  movel([0.337067, -0.792207, -2.792280, -1.127903, 1.570796, 1.907863],accel_mss,speed_ms,0,blend_radius_m)
  movel([0.336030, -0.792065, -2.792303, -1.128021, 1.570796, 1.906826],accel_mss,speed_ms,0,blend_radius_m)
  movel([0.330509, -0.790300, -2.792596, -1.129493, 1.570796, 1.901306],accel_mss,speed_ms,0,blend_radius_m)
  movel([0.325271, -0.788116, -2.792957, -1.131316, 1.570796, 1.896067],accel_mss,speed_ms,0,blend_radius_m)
  movel([0.320318, -0.785517, -2.793383, -1.133490, 1.570796, 1.891115],accel_mss,speed_ms,0,blend_radius_m)
  movel([0.315671, -0.782494, -2.793873, -1.136022, 1.570796, 1.886468],accel_mss,speed_ms,0,blend_radius_m)
  movel([0.314088, -0.781197, -2.794083, -1.137109, 1.570796, 1.884885],accel_mss,speed_ms,0,blend_radius_m)
  movel([0.312919, -0.779429, -2.794366, -1.138594, 1.570796, 1.883716],accel_mss,speed_ms,0,blend_radius_m)
  movel([0.312565, -0.778043, -2.794588, -1.139758, 1.570796, 1.883362],accel_mss,speed_ms,0,blend_radius_m)
  movel([0.312427, -0.776467, -2.794838, -1.141084, 1.570796, 1.883224],accel_mss,speed_ms,0,blend_radius_m)
  movel([0.312533, -0.772984, -2.795388, -1.144017, 1.570796, 1.883329],accel_mss,speed_ms,0,blend_radius_m)
  movel([0.314201, -0.759545, -2.797451, -1.155393, 1.570796, 1.884998],accel_mss,speed_ms,0,blend_radius_m)
  movel([0.314322, -0.755972, -2.797984, -1.158433, 1.570796, 1.885118],accel_mss,speed_ms,0,blend_radius_m)
  movel([0.313995, -0.753066, -2.798414, -1.160909, 1.570796, 1.884791],accel_mss,speed_ms,0,blend_radius_m)
  movel([0.313608, -0.751988, -2.798572, -1.161829, 1.570796, 1.884404],accel_mss,speed_ms,0,blend_radius_m)
  movel([0.313044, -0.751216, -2.798685, -1.162488, 1.570796, 1.883841],accel_mss,speed_ms,0,blend_radius_m)
  movel([0.312284, -0.750809, -2.798744, -1.162836, 1.570796, 1.883080],accel_mss,speed_ms,0,blend_radius_m)
  movel([0.311307, -0.750804, -2.798745, -1.162840, 1.570796, 1.882104],accel_mss,speed_ms,0,blend_radius_m)
  movel([0.309324, -0.751441, -2.798652, -1.162296, 1.570796, 1.880120],accel_mss,speed_ms,0,blend_radius_m)
  movel([0.308425, -0.751616, -2.798626, -1.162147, 1.570796, 1.879221],accel_mss,speed_ms,0,blend_radius_m)
  movel([0.307786, -0.751386, -2.798660, -1.162343, 1.570796, 1.878582],accel_mss,speed_ms,0,blend_radius_m)
  movel([0.307584, -0.750201, -2.798833, -1.163355, 1.570796, 1.878380],accel_mss,speed_ms,0,blend_radius_m)
  movel([0.307977, -0.748520, -2.799077, -1.164791, 1.570796, 1.878773],accel_mss,speed_ms,0,blend_radius_m)
  movel([0.309463, -0.743009, -2.799868, -1.169512, 1.570796, 1.880260],accel_mss,speed_ms,0,blend_radius_m)
  movel([0.310630, -0.737685, -2.800619, -1.174085, 1.570796, 1.881426],accel_mss,speed_ms,0,blend_radius_m)
  movel([0.312165, -0.727491, -2.802019, -1.182879, 1.570796, 1.882961],accel_mss,speed_ms,0,blend_radius_m)
  movel([0.312944, -0.717680, -2.803320, -1.191389, 1.570796, 1.883740],accel_mss,speed_ms,0,blend_radius_m)
  movel([0.313326, -0.707992, -2.804562, -1.199834, 1.570796, 1.884122],accel_mss,speed_ms,0,blend_radius_m)
  speed_ms = 0.005
  movel([0.313326, -0.701025, -2.797945, -1.213418, 1.570796, 1.884122],accel_mss,speed_ms,0,blend_radius_m)
  speed_ms = 0.040
  movel([0.305588, -0.719229, -2.795588, -1.197572, 1.570796, 1.876385],accel_mss,speed_ms,0,blend_radius_m)
  speed_ms = 0.005
  movel([0.305588, -0.726439, -2.802160, -1.183790, 1.570796, 1.876385],accel_mss,speed_ms,0,blend_radius_m)
  speed_ms = 0.025
  movel([0.301170, -0.738509, -2.800504, -1.173377, 1.570796, 1.871966],accel_mss,speed_ms,0,blend_radius_m)
  movel([0.298692, -0.744594, -2.799642, -1.168153, 1.570796, 1.869489],accel_mss,speed_ms,0,blend_radius_m)
  movel([0.296052, -0.750689, -2.798762, -1.162938, 1.570796, 1.866849],accel_mss,speed_ms,0,blend_radius_m)
  movel([0.293909, -0.749383, -2.798952, -1.164054, 1.570796, 1.864706],accel_mss,speed_ms,0,blend_radius_m)
  movel([0.293492, -0.749233, -2.798974, -1.164182, 1.570796, 1.864289],accel_mss,speed_ms,0,blend_radius_m)
  movel([0.292925, -0.749435, -2.798944, -1.164009, 1.570796, 1.863721],accel_mss,speed_ms,0,blend_radius_m)
  movel([0.292315, -0.750102, -2.798847, -1.163439, 1.570796, 1.863111],accel_mss,speed_ms,0,blend_radius_m)
  movel([0.291839, -0.750915, -2.798729, -1.162745, 1.570796, 1.862635],accel_mss,speed_ms,0,blend_radius_m)
  movel([0.288894, -0.755925, -2.797991, -1.158473, 1.570796, 1.859691],accel_mss,speed_ms,0,blend_radius_m)
  movel([0.285493, -0.760805, -2.797261, -1.154323, 1.570796, 1.856290],accel_mss,speed_ms,0,blend_radius_m)
  movel([0.284595, -0.761864, -2.797101, -1.153424, 1.570796, 1.855391],accel_mss,speed_ms,0,blend_radius_m)
  movel([0.283710, -0.762451, -2.797012, -1.152926, 1.570796, 1.854506],accel_mss,speed_ms,0,blend_radius_m)
  movel([0.283279, -0.762203, -2.797050, -1.153136, 1.570796, 1.854075],accel_mss,speed_ms,0,blend_radius_m)
  movel([0.283199, -0.761526, -2.797152, -1.153711, 1.570796, 1.853995],accel_mss,speed_ms,0,blend_radius_m)
  movel([0.283611, -0.756734, -2.797871, -1.157784, 1.570796, 1.854408],accel_mss,speed_ms,0,blend_radius_m)
  movel([0.284807, -0.751427, -2.798654, -1.162308, 1.570796, 1.855604],accel_mss,speed_ms,0,blend_radius_m)
  speed_ms = 0.005
  movel([0.284807, -0.743907, -2.792145, -1.176337, 1.570796, 1.855604],accel_mss,speed_ms,0,blend_radius_m)
  speed_ms = 0.040
  movel([0.290706, -0.750918, -2.791114, -1.170358, 1.570796, 1.861503],accel_mss,speed_ms,0,blend_radius_m)
  speed_ms = 0.005
  movel([0.290706, -0.758522, -2.797604, -1.156263, 1.570796, 1.861503],accel_mss,speed_ms,0,blend_radius_m)
  speed_ms = 0.025
  movel([0.289009, -0.766268, -2.796430, -1.149691, 1.570796, 1.859805],accel_mss,speed_ms,0,blend_radius_m)
  movel([0.287811, -0.770306, -2.795806, -1.146277, 1.570796, 1.858608],accel_mss,speed_ms,0,blend_radius_m)
  movel([0.284778, -0.778595, -2.794500, -1.139294, 1.570796, 1.855575],accel_mss,speed_ms,0,blend_radius_m)
  movel([0.282956, -0.782810, -2.793822, -1.135757, 1.570796, 1.853753],accel_mss,speed_ms,0,blend_radius_m)
  movel([0.278747, -0.791286, -2.792433, -1.128671, 1.570796, 1.849544],accel_mss,speed_ms,0,blend_radius_m)
  movel([0.279478, -0.788663, -2.792867, -1.130860, 1.570796, 1.850275],accel_mss,speed_ms,0,blend_radius_m)
  movel([0.279565, -0.786419, -2.793235, -1.132735, 1.570796, 1.850361],accel_mss,speed_ms,0,blend_radius_m)
  movel([0.279016, -0.784705, -2.793515, -1.134169, 1.570796, 1.849813],accel_mss,speed_ms,0,blend_radius_m)
  movel([0.277841, -0.783676, -2.793682, -1.135031, 1.570796, 1.848637],accel_mss,speed_ms,0,blend_radius_m)
  speed_ms = 0.005
  movel([0.277841, -0.775786, -2.787260, -1.149343, 1.570796, 1.848637],accel_mss,speed_ms,0,blend_radius_m)
  speed_ms = 0.040
  movel([0.251919, -0.792770, -2.784449, -1.135169, 1.570796, 1.822716],accel_mss,speed_ms,0,blend_radius_m)
  speed_ms = 0.005
  movel([0.251919, -0.800843, -2.790822, -1.120725, 1.570796, 1.822716],accel_mss,speed_ms,0,blend_radius_m)
  speed_ms = 0.025
  movel([0.247378, -0.806648, -2.789820, -1.115921, 1.570796, 1.818174],accel_mss,speed_ms,0,blend_radius_m)
  movel([0.242549, -0.812092, -2.788864, -1.111433, 1.570796, 1.813345],accel_mss,speed_ms,0,blend_radius_m)
  movel([0.237519, -0.817097, -2.787971, -1.107321, 1.570796, 1.808315],accel_mss,speed_ms,0,blend_radius_m)
  movel([0.232368, -0.821580, -2.787160, -1.103649, 1.570796, 1.803164],accel_mss,speed_ms,0,blend_radius_m)
  movel([0.233688, -0.818996, -2.787629, -1.105764, 1.570796, 1.804484],accel_mss,speed_ms,0,blend_radius_m)
  movel([0.234683, -0.816593, -2.788062, -1.107734, 1.570796, 1.805479],accel_mss,speed_ms,0,blend_radius_m)
  movel([0.235280, -0.814585, -2.788421, -1.109383, 1.570796, 1.806076],accel_mss,speed_ms,0,blend_radius_m)
  movel([0.235407, -0.813183, -2.788670, -1.110536, 1.570796, 1.806203],accel_mss,speed_ms,0,blend_radius_m)
  movel([0.234984, -0.812617, -2.788771, -1.111001, 1.570796, 1.805780],accel_mss,speed_ms,0,blend_radius_m)
  movel([0.234547, -0.812711, -2.788754, -1.110924, 1.570796, 1.805344],accel_mss,speed_ms,0,blend_radius_m)
  movel([0.233940, -0.813094, -2.788686, -1.110609, 1.570796, 1.804736],accel_mss,speed_ms,0,blend_radius_m)
  movel([0.232209, -0.814833, -2.788377, -1.109180, 1.570796, 1.803005],accel_mss,speed_ms,0,blend_radius_m)
  movel([0.227802, -0.820578, -2.787342, -1.104469, 1.570796, 1.798598],accel_mss,speed_ms,0,blend_radius_m)
  movel([0.225752, -0.823067, -2.786889, -1.102433, 1.570796, 1.796549],accel_mss,speed_ms,0,blend_radius_m)
  movel([0.221376, -0.827745, -2.786027, -1.098617, 1.570796, 1.792172],accel_mss,speed_ms,0,blend_radius_m)
  movel([0.219102, -0.829874, -2.785631, -1.096884, 1.570796, 1.789898],accel_mss,speed_ms,0,blend_radius_m)
  movel([0.216804, -0.831814, -2.785268, -1.095307, 1.570796, 1.787600],accel_mss,speed_ms,0,blend_radius_m)
  movel([0.214506, -0.833546, -2.784942, -1.093901, 1.570796, 1.785302],accel_mss,speed_ms,0,blend_radius_m)
  movel([0.212240, -0.835024, -2.784662, -1.092702, 1.570796, 1.783037],accel_mss,speed_ms,0,blend_radius_m)
  movel([0.215104, -0.830931, -2.785433, -1.096025, 1.570796, 1.785901],accel_mss,speed_ms,0,blend_radius_m)
  movel([0.217906, -0.826781, -2.786206, -1.099402, 1.570796, 1.788702],accel_mss,speed_ms,0,blend_radius_m)
  movel([0.219209, -0.824080, -2.786703, -1.101606, 1.570796, 1.790005],accel_mss,speed_ms,0,blend_radius_m)
  movel([0.219966, -0.821533, -2.787169, -1.103687, 1.570796, 1.790763],accel_mss,speed_ms,0,blend_radius_m)
  movel([0.219920, -0.820731, -2.787315, -1.104343, 1.570796, 1.790716],accel_mss,speed_ms,0,blend_radius_m)
  movel([0.219466, -0.820469, -2.787362, -1.104558, 1.570796, 1.790262],accel_mss,speed_ms,0,blend_radius_m)
  movel([0.218525, -0.820910, -2.787282, -1.104197, 1.570796, 1.789321],accel_mss,speed_ms,0,blend_radius_m)
  movel([0.217006, -0.822224, -2.787043, -1.103122, 1.570796, 1.787803],accel_mss,speed_ms,0,blend_radius_m)
  movel([0.209003, -0.830286, -2.785554, -1.096549, 1.570796, 1.779799],accel_mss,speed_ms,0,blend_radius_m)
  movel([0.205006, -0.833828, -2.784889, -1.093672, 1.570796, 1.775803],accel_mss,speed_ms,0,blend_radius_m)
  movel([0.203015, -0.835288, -2.784612, -1.092488, 1.570796, 1.773811],accel_mss,speed_ms,0,blend_radius_m)
  movel([0.201023, -0.836475, -2.784387, -1.091527, 1.570796, 1.771819],accel_mss,speed_ms,0,blend_radius_m)
  speed_ms = 0.005
  movel([0.201023, -0.828056, -2.778123, -1.106210, 1.570796, 1.771819],accel_mss,speed_ms,0,blend_radius_m)
  speed_ms = 0.040
  movel([0.238662, -0.773617, -2.787609, -1.151163, 1.570796, 1.809458],accel_mss,speed_ms,0,blend_radius_m)
  speed_ms = 0.005
  movel([0.238662, -0.781483, -2.794037, -1.136870, 1.570796, 1.809458],accel_mss,speed_ms,0,blend_radius_m)
  speed_ms = 0.025
  movel([0.238890, -0.778419, -2.794528, -1.139442, 1.570796, 1.809686],accel_mss,speed_ms,0,blend_radius_m)
  movel([0.239732, -0.775008, -2.795069, -1.142312, 1.570796, 1.810528],accel_mss,speed_ms,0,blend_radius_m)
  movel([0.241121, -0.771324, -2.795647, -1.145418, 1.570796, 1.811917],accel_mss,speed_ms,0,blend_radius_m)
  movel([0.242984, -0.767463, -2.796246, -1.148680, 1.570796, 1.813781],accel_mss,speed_ms,0,blend_radius_m)
  movel([0.245268, -0.763496, -2.796853, -1.152040, 1.570796, 1.816064],accel_mss,speed_ms,0,blend_radius_m)
  movel([0.247890, -0.759528, -2.797453, -1.155408, 1.570796, 1.818687],accel_mss,speed_ms,0,blend_radius_m)
  movel([0.250794, -0.755633, -2.798035, -1.158721, 1.570796, 1.821590],accel_mss,speed_ms,0,blend_radius_m)
  movel([0.253896, -0.751916, -2.798582, -1.161891, 1.570796, 1.824692],accel_mss,speed_ms,0,blend_radius_m)
  movel([0.257898, -0.747597, -2.799211, -1.165581, 1.570796, 1.828695],accel_mss,speed_ms,0,blend_radius_m)
  movel([0.266086, -0.739112, -2.800419, -1.172858, 1.570796, 1.836882],accel_mss,speed_ms,0,blend_radius_m)
  movel([0.270058, -0.734609, -2.801046, -1.176734, 1.570796, 1.840855],accel_mss,speed_ms,0,blend_radius_m)
  movel([0.273771, -0.729657, -2.801725, -1.181007, 1.570796, 1.844568],accel_mss,speed_ms,0,blend_radius_m)
  movel([0.275420, -0.727072, -2.802075, -1.183242, 1.570796, 1.846216],accel_mss,speed_ms,0,blend_radius_m)
  movel([0.276854, -0.724500, -2.802420, -1.185469, 1.570796, 1.847650],accel_mss,speed_ms,0,blend_radius_m)
  movel([0.278016, -0.722006, -2.802752, -1.187631, 1.570796, 1.848812],accel_mss,speed_ms,0,blend_radius_m)
  movel([0.278854, -0.719652, -2.803062, -1.189675, 1.570796, 1.849650],accel_mss,speed_ms,0,blend_radius_m)
  movel([0.279296, -0.717519, -2.803341, -1.191528, 1.570796, 1.850092],accel_mss,speed_ms,0,blend_radius_m)
  movel([0.279283, -0.715676, -2.803581, -1.193133, 1.570796, 1.850080],accel_mss,speed_ms,0,blend_radius_m)
  speed_ms = 0.005
  movel([0.279283, -0.708606, -2.796982, -1.206801, 1.570796, 1.850080],accel_mss,speed_ms,0,blend_radius_m)
  speed_ms = 0.040
  movel([0.278218, -0.694550, -2.798748, -1.219091, 1.570796, 1.849015],accel_mss,speed_ms,0,blend_radius_m)
  speed_ms = 0.005
  movel([0.278218, -0.701428, -2.805380, -1.205581, 1.570796, 1.849015],accel_mss,speed_ms,0,blend_radius_m)
  speed_ms = 0.025
  movel([0.274128, -0.714706, -2.803706, -1.193977, 1.570796, 1.844925],accel_mss,speed_ms,0,blend_radius_m)
  movel([0.272708, -0.717821, -2.803302, -1.191267, 1.570796, 1.843504],accel_mss,speed_ms,0,blend_radius_m)
  movel([0.270637, -0.720929, -2.802894, -1.188566, 1.570796, 1.841433],accel_mss,speed_ms,0,blend_radius_m)
  movel([0.268156, -0.723829, -2.802510, -1.186050, 1.570796, 1.838952],accel_mss,speed_ms,0,blend_radius_m)
  movel([0.259858, -0.732396, -2.801351, -1.178642, 1.570796, 1.830654],accel_mss,speed_ms,0,blend_radius_m)
  movel([0.257055, -0.735659, -2.800901, -1.175829, 1.570796, 1.827852],accel_mss,speed_ms,0,blend_radius_m)
  movel([0.254399, -0.739041, -2.800429, -1.172919, 1.570796, 1.825196],accel_mss,speed_ms,0,blend_radius_m)
  movel([0.251913, -0.742499, -2.799941, -1.169949, 1.570796, 1.822709],accel_mss,speed_ms,0,blend_radius_m)
  movel([0.249806, -0.745929, -2.799451, -1.167009, 1.570796, 1.820602],accel_mss,speed_ms,0,blend_radius_m)
  movel([0.248006, -0.749350, -2.798957, -1.164082, 1.570796, 1.818802],accel_mss,speed_ms,0,blend_radius_m)
  movel([0.246241, -0.752742, -2.798461, -1.161185, 1.570796, 1.817038],accel_mss,speed_ms,0,blend_radius_m)
  movel([0.244246, -0.756094, -2.797966, -1.158329, 1.570796, 1.815042],accel_mss,speed_ms,0,blend_radius_m)
  movel([0.242758, -0.750446, -2.798797, -1.163146, 1.570796, 1.813555],accel_mss,speed_ms,0,blend_radius_m)
  movel([0.243050, -0.748448, -2.799088, -1.164853, 1.570796, 1.813846],accel_mss,speed_ms,0,blend_radius_m)
  movel([0.243651, -0.746324, -2.799394, -1.166671, 1.570796, 1.814448],accel_mss,speed_ms,0,blend_radius_m)
  movel([0.244562, -0.744068, -2.799717, -1.168603, 1.570796, 1.815359],accel_mss,speed_ms,0,blend_radius_m)
  movel([0.245801, -0.741661, -2.800060, -1.170669, 1.570796, 1.816598],accel_mss,speed_ms,0,blend_radius_m)
  movel([0.248098, -0.738282, -2.800535, -1.173572, 1.570796, 1.818894],accel_mss,speed_ms,0,blend_radius_m)
  movel([0.251441, -0.734149, -2.801110, -1.177130, 1.570796, 1.822238],accel_mss,speed_ms,0,blend_radius_m)
  movel([0.259675, -0.724773, -2.802384, -1.185232, 1.570796, 1.830471],accel_mss,speed_ms,0,blend_radius_m)
  movel([0.263755, -0.720127, -2.803000, -1.189262, 1.570796, 1.834551],accel_mss,speed_ms,0,blend_radius_m)
  movel([0.267253, -0.715908, -2.803551, -1.192931, 1.570796, 1.838049],accel_mss,speed_ms,0,blend_radius_m)
  movel([0.269743, -0.712436, -2.803998, -1.195955, 1.570796, 1.840539],accel_mss,speed_ms,0,blend_radius_m)
  movel([0.270479, -0.711072, -2.804172, -1.197145, 1.570796, 1.841275],accel_mss,speed_ms,0,blend_radius_m)
  movel([0.270799, -0.710010, -2.804307, -1.198072, 1.570796, 1.841595],accel_mss,speed_ms,0,blend_radius_m)
  speed_ms = 0.005
  movel([0.270799, -0.703016, -2.797695, -1.211678, 1.570796, 1.841595],accel_mss,speed_ms,0,blend_radius_m)
  speed_ms = 0.040
  movel([0.256086, -0.705862, -2.797334, -1.209193, 1.570796, 1.826882],accel_mss,speed_ms,0,blend_radius_m)
  speed_ms = 0.005
  movel([0.256086, -0.712894, -2.803939, -1.195555, 1.570796, 1.826882],accel_mss,speed_ms,0,blend_radius_m)
  speed_ms = 0.025
  movel([0.254666, -0.713145, -2.803907, -1.195337, 1.570796, 1.825462],accel_mss,speed_ms,0,blend_radius_m)
  movel([0.253508, -0.712972, -2.803929, -1.195488, 1.570796, 1.824304],accel_mss,speed_ms,0,blend_radius_m)
  movel([0.251855, -0.711627, -2.804101, -1.196661, 1.570796, 1.822651],accel_mss,speed_ms,0,blend_radius_m)
  movel([0.250882, -0.709349, -2.804391, -1.198649, 1.570796, 1.821679],accel_mss,speed_ms,0,blend_radius_m)
  movel([0.250362, -0.706617, -2.804735, -1.201037, 1.570796, 1.821158],accel_mss,speed_ms,0,blend_radius_m)
  movel([0.250376, -0.705463, -2.804880, -1.202047, 1.570796, 1.821172],accel_mss,speed_ms,0,blend_radius_m)
  movel([0.251431, -0.703143, -2.805168, -1.204078, 1.570796, 1.822227],accel_mss,speed_ms,0,blend_radius_m)
  movel([0.255097, -0.696419, -2.805991, -1.209980, 1.570796, 1.825893],accel_mss,speed_ms,0,blend_radius_m)
  movel([0.261993, -0.682881, -2.807586, -1.221922, 1.570796, 1.832789],accel_mss,speed_ms,0,blend_radius_m)
  movel([0.265206, -0.676101, -2.808355, -1.227933, 1.570796, 1.836002],accel_mss,speed_ms,0,blend_radius_m)
  speed_ms = 0.005
  movel([0.265206, -0.669577, -2.801667, -1.241144, 1.570796, 1.836002],accel_mss,speed_ms,0,blend_radius_m)
  speed_ms = 0.040
  movel([0.255172, -0.676970, -2.800832, -1.234588, 1.570796, 1.825968],accel_mss,speed_ms,0,blend_radius_m)
  speed_ms = 0.005
  movel([0.255172, -0.683600, -2.807503, -1.221285, 1.570796, 1.825968],accel_mss,speed_ms,0,blend_radius_m)
  speed_ms = 0.025
  movel([0.253576, -0.687576, -2.807042, -1.217771, 1.570796, 1.824373],accel_mss,speed_ms,0,blend_radius_m)
  movel([0.251612, -0.691649, -2.806562, -1.214178, 1.570796, 1.822409],accel_mss,speed_ms,0,blend_radius_m)
  movel([0.249200, -0.695639, -2.806085, -1.210665, 1.570796, 1.819996],accel_mss,speed_ms,0,blend_radius_m)
  movel([0.247798, -0.697558, -2.805853, -1.208978, 1.570796, 1.818594],accel_mss,speed_ms,0,blend_radius_m)
  movel([0.244762, -0.701197, -2.805408, -1.205783, 1.570796, 1.815558],accel_mss,speed_ms,0,blend_radius_m)
  movel([0.243999, -0.702815, -2.805209, -1.204365, 1.570796, 1.814795],accel_mss,speed_ms,0,blend_radius_m)
  movel([0.239388, -0.714876, -2.803684, -1.193828, 1.570796, 1.810184],accel_mss,speed_ms,0,blend_radius_m)
  movel([0.238976, -0.716027, -2.803535, -1.192826, 1.570796, 1.809772],accel_mss,speed_ms,0,blend_radius_m)
  movel([0.238840, -0.717001, -2.803409, -1.191979, 1.570796, 1.809637],accel_mss,speed_ms,0,blend_radius_m)
  movel([0.239436, -0.717697, -2.803318, -1.191374, 1.570796, 1.810232],accel_mss,speed_ms,0,blend_radius_m)
  movel([0.240542, -0.717756, -2.803310, -1.191323, 1.570796, 1.811338],accel_mss,speed_ms,0,blend_radius_m)
  movel([0.243805, -0.717753, -2.803311, -1.191325, 1.570796, 1.814601],accel_mss,speed_ms,0,blend_radius_m)
  movel([0.246751, -0.718260, -2.803245, -1.190885, 1.570796, 1.817547],accel_mss,speed_ms,0,blend_radius_m)
  movel([0.249147, -0.719502, -2.803082, -1.189805, 1.570796, 1.819943],accel_mss,speed_ms,0,blend_radius_m)
  movel([0.250740, -0.721722, -2.802789, -1.187877, 1.570796, 1.821537],accel_mss,speed_ms,0,blend_radius_m)
  speed_ms = 0.005
  movel([0.250740, -0.714574, -2.796205, -1.201610, 1.570796, 1.821537],accel_mss,speed_ms,0,blend_radius_m)
  speed_ms = 0.040
  movel([0.239180, -0.744721, -2.792026, -1.175642, 1.570796, 1.809976],accel_mss,speed_ms,0,blend_radius_m)
  speed_ms = 0.005
  movel([0.239180, -0.752251, -2.798533, -1.161605, 1.570796, 1.809976],accel_mss,speed_ms,0,blend_radius_m)
  speed_ms = 0.025
  movel([0.238467, -0.752976, -2.798427, -1.160986, 1.570796, 1.809264],accel_mss,speed_ms,0,blend_radius_m)
  movel([0.237810, -0.753876, -2.798294, -1.160218, 1.570796, 1.808607],accel_mss,speed_ms,0,blend_radius_m)
  movel([0.235162, -0.758478, -2.797611, -1.156301, 1.570796, 1.805958],accel_mss,speed_ms,0,blend_radius_m)
  movel([0.234732, -0.758919, -2.797545, -1.155925, 1.570796, 1.805529],accel_mss,speed_ms,0,blend_radius_m)
  movel([0.234120, -0.759144, -2.797511, -1.155734, 1.570796, 1.804916],accel_mss,speed_ms,0,blend_radius_m)
  movel([0.233671, -0.758910, -2.797546, -1.155933, 1.570796, 1.804467],accel_mss,speed_ms,0,blend_radius_m)
  movel([0.233188, -0.757524, -2.797753, -1.157112, 1.570796, 1.803984],accel_mss,speed_ms,0,blend_radius_m)
  movel([0.233194, -0.754285, -2.798234, -1.159870, 1.570796, 1.803991],accel_mss,speed_ms,0,blend_radius_m)
  movel([0.234136, -0.750704, -2.798760, -1.162926, 1.570796, 1.804933],accel_mss,speed_ms,0,blend_radius_m)
  movel([0.235569, -0.746865, -2.799316, -1.166208, 1.570796, 1.806365],accel_mss,speed_ms,0,blend_radius_m)
  movel([0.237248, -0.742984, -2.799872, -1.169533, 1.570796, 1.808045],accel_mss,speed_ms,0,blend_radius_m)
  movel([0.239202, -0.739157, -2.800413, -1.172820, 1.570796, 1.809999],accel_mss,speed_ms,0,blend_radius_m)
  movel([0.241419, -0.735387, -2.800939, -1.176063, 1.570796, 1.812215],accel_mss,speed_ms,0,blend_radius_m)
  movel([0.243887, -0.731674, -2.801450, -1.179265, 1.570796, 1.814683],accel_mss,speed_ms,0,blend_radius_m)
  movel([0.246599, -0.728014, -2.801948, -1.182427, 1.570796, 1.817396],accel_mss,speed_ms,0,blend_radius_m)
  movel([0.249538, -0.724415, -2.802431, -1.185542, 1.570796, 1.820334],accel_mss,speed_ms,0,blend_radius_m)
  movel([0.252702, -0.720865, -2.802902, -1.188621, 1.570796, 1.823499],accel_mss,speed_ms,0,blend_radius_m)
  movel([0.256073, -0.717373, -2.803360, -1.191656, 1.570796, 1.826870],accel_mss,speed_ms,0,blend_radius_m)
  movel([0.260755, -0.712155, -2.804034, -1.196200, 1.570796, 1.831551],accel_mss,speed_ms,0,blend_radius_m)
  movel([0.265685, -0.706033, -2.804808, -1.201548, 1.570796, 1.836482],accel_mss,speed_ms,0,blend_radius_m)
  movel([0.271037, -0.698934, -2.805685, -1.207769, 1.570796, 1.841833],accel_mss,speed_ms,0,blend_radius_m)
  speed_ms = 0.005
  movel([0.271037, -0.692090, -2.799048, -1.221251, 1.570796, 1.841833],accel_mss,speed_ms,0,blend_radius_m)
  speed_ms = 0.040
  movel([0.266633, -0.693684, -2.798854, -1.219851, 1.570796, 1.837429],accel_mss,speed_ms,0,blend_radius_m)
  speed_ms = 0.005
  movel([0.266633, -0.700551, -2.805488, -1.206351, 1.570796, 1.837429],accel_mss,speed_ms,0,blend_radius_m)
  speed_ms = 0.025
  movel([0.271058, -0.690929, -2.806647, -1.214812, 1.570796, 1.841854],accel_mss,speed_ms,0,blend_radius_m)
  movel([0.275991, -0.681101, -2.807790, -1.223498, 1.570796, 1.846787],accel_mss,speed_ms,0,blend_radius_m)
  movel([0.278750, -0.676151, -2.808350, -1.227888, 1.570796, 1.849546],accel_mss,speed_ms,0,blend_radius_m)
  movel([0.281743, -0.671202, -2.808898, -1.232288, 1.570796, 1.852540],accel_mss,speed_ms,0,blend_radius_m)
  movel([0.285025, -0.666265, -2.809436, -1.236688, 1.570796, 1.855822],accel_mss,speed_ms,0,blend_radius_m)
  movel([0.288616, -0.661374, -2.809958, -1.241057, 1.570796, 1.859412],accel_mss,speed_ms,0,blend_radius_m)
  movel([0.298570, -0.649107, -2.811222, -1.252060, 1.570796, 1.869366],accel_mss,speed_ms,0,blend_radius_m)
  movel([0.302903, -0.643471, -2.811782, -1.257136, 1.570796, 1.873699],accel_mss,speed_ms,0,blend_radius_m)
  movel([0.304959, -0.640578, -2.812065, -1.259747, 1.570796, 1.875755],accel_mss,speed_ms,0,blend_radius_m)
  movel([0.306841, -0.637624, -2.812349, -1.262415, 1.570796, 1.877638],accel_mss,speed_ms,0,blend_radius_m)
  movel([0.311183, -0.628769, -2.813182, -1.270439, 1.570796, 1.881979],accel_mss,speed_ms,0,blend_radius_m)
  speed_ms = 0.005
  movel([0.311183, -0.622959, -2.806401, -1.283029, 1.570796, 1.881979],accel_mss,speed_ms,0,blend_radius_m)
  speed_ms = 0.040
  movel([0.321759, -0.602546, -2.808192, -1.301652, 1.570796, 1.892555],accel_mss,speed_ms,0,blend_radius_m)
  speed_ms = 0.005
  movel([0.321759, -0.608023, -2.815008, -1.289358, 1.570796, 1.892555],accel_mss,speed_ms,0,blend_radius_m)
  speed_ms = 0.025
  movel([0.325188, -0.600693, -2.815612, -1.296084, 1.570796, 1.895984],accel_mss,speed_ms,0,blend_radius_m)
  movel([0.327388, -0.596990, -2.815910, -1.299490, 1.570796, 1.898185],accel_mss,speed_ms,0,blend_radius_m)
  movel([0.330084, -0.593376, -2.816195, -1.302818, 1.570796, 1.900880],accel_mss,speed_ms,0,blend_radius_m)
  movel([0.332238, -0.591038, -2.816376, -1.304975, 1.570796, 1.903034],accel_mss,speed_ms,0,blend_radius_m)
  movel([0.334479, -0.588925, -2.816539, -1.306925, 1.570796, 1.905275],accel_mss,speed_ms,0,blend_radius_m)
  movel([0.339064, -0.585048, -2.816832, -1.310509, 1.570796, 1.909861],accel_mss,speed_ms,0,blend_radius_m)
  movel([0.343198, -0.581242, -2.817115, -1.314032, 1.570796, 1.913994],accel_mss,speed_ms,0,blend_radius_m)
  movel([0.346574, -0.577426, -2.817392, -1.317571, 1.570796, 1.917370],accel_mss,speed_ms,0,blend_radius_m)
  movel([0.353165, -0.568512, -2.818019, -1.325858, 1.570796, 1.923961],accel_mss,speed_ms,0,blend_radius_m)
  movel([0.354587, -0.566740, -2.818140, -1.327509, 1.570796, 1.925383],accel_mss,speed_ms,0,blend_radius_m)
  movel([0.356113, -0.565141, -2.818248, -1.329000, 1.570796, 1.926909],accel_mss,speed_ms,0,blend_radius_m)
  movel([0.359378, -0.562332, -2.818436, -1.331621, 1.570796, 1.930174],accel_mss,speed_ms,0,blend_radius_m)
  movel([0.365995, -0.557274, -2.818767, -1.336348, 1.570796, 1.936792],accel_mss,speed_ms,0,blend_radius_m)
  movel([0.373073, -0.551234, -2.819149, -1.342006, 1.570796, 1.943869],accel_mss,speed_ms,0,blend_radius_m)
  movel([0.376615, -0.547904, -2.819354, -1.345131, 1.570796, 1.947411],accel_mss,speed_ms,0,blend_radius_m)
  movel([0.380090, -0.544218, -2.819576, -1.348595, 1.570796, 1.950886],accel_mss,speed_ms,0,blend_radius_m)
  movel([0.382697, -0.540897, -2.819772, -1.351720, 1.570796, 1.953493],accel_mss,speed_ms,0,blend_radius_m)
  movel([0.384821, -0.537477, -2.819969, -1.354943, 1.570796, 1.955617],accel_mss,speed_ms,0,blend_radius_m)
  movel([0.385968, -0.534592, -2.820132, -1.357665, 1.570796, 1.956764],accel_mss,speed_ms,0,blend_radius_m)
  movel([0.386018, -0.533554, -2.820190, -1.358645, 1.570796, 1.956814],accel_mss,speed_ms,0,blend_radius_m)
  movel([0.385633, -0.532896, -2.820226, -1.359267, 1.570796, 1.956430],accel_mss,speed_ms,0,blend_radius_m)
  movel([0.384024, -0.532480, -2.820249, -1.359660, 1.570796, 1.954820],accel_mss,speed_ms,0,blend_radius_m)
  movel([0.381703, -0.532851, -2.820229, -1.359309, 1.570796, 1.952500],accel_mss,speed_ms,0,blend_radius_m)
  movel([0.378837, -0.533912, -2.820170, -1.358307, 1.570796, 1.949633],accel_mss,speed_ms,0,blend_radius_m)
  movel([0.375629, -0.535524, -2.820080, -1.356785, 1.570796, 1.946425],accel_mss,speed_ms,0,blend_radius_m)
  movel([0.372254, -0.537591, -2.819962, -1.354836, 1.570796, 1.943051],accel_mss,speed_ms,0,blend_radius_m)
  movel([0.368906, -0.539977, -2.819825, -1.352587, 1.570796, 1.939702],accel_mss,speed_ms,0,blend_radius_m)
  movel([0.365765, -0.542576, -2.819673, -1.350140, 1.570796, 1.936562],accel_mss,speed_ms,0,blend_radius_m)
  movel([0.363011, -0.545269, -2.819513, -1.347607, 1.570796, 1.933807],accel_mss,speed_ms,0,blend_radius_m)
  movel([0.359228, -0.549801, -2.819237, -1.343350, 1.570796, 1.930024],accel_mss,speed_ms,0,blend_radius_m)
  movel([0.348676, -0.563729, -2.818343, -1.330317, 1.570796, 1.919472],accel_mss,speed_ms,0,blend_radius_m)
  movel([0.341420, -0.572642, -2.817732, -1.322014, 1.570796, 1.912216],accel_mss,speed_ms,0,blend_radius_m)
  movel([0.334837, -0.579815, -2.817219, -1.315355, 1.570796, 1.905633],accel_mss,speed_ms,0,blend_radius_m)
  movel([0.331585, -0.583292, -2.816963, -1.312134, 1.570796, 1.902381],accel_mss,speed_ms,0,blend_radius_m)
  movel([0.328499, -0.586903, -2.816693, -1.308793, 1.570796, 1.899296],accel_mss,speed_ms,0,blend_radius_m)
  movel([0.325566, -0.590822, -2.816393, -1.305174, 1.570796, 1.896362],accel_mss,speed_ms,0,blend_radius_m)
  movel([0.322921, -0.594763, -2.816086, -1.301540, 1.570796, 1.893717],accel_mss,speed_ms,0,blend_radius_m)
  movel([0.320533, -0.598711, -2.815772, -1.297905, 1.570796, 1.891330],accel_mss,speed_ms,0,blend_radius_m)
  movel([0.318373, -0.602637, -2.815454, -1.294298, 1.570796, 1.889170],accel_mss,speed_ms,0,blend_radius_m)
  movel([0.314600, -0.610358, -2.814811, -1.287220, 1.570796, 1.885397],accel_mss,speed_ms,0,blend_radius_m)
  movel([0.311326, -0.617785, -2.814170, -1.280434, 1.570796, 1.882122],accel_mss,speed_ms,0,blend_radius_m)
  speed_ms = 0.005
  movel([0.311326, -0.612149, -2.807370, -1.292869, 1.570796, 1.882122],accel_mss,speed_ms,0,blend_radius_m)
  speed_ms = 0.040
  movel([0.303174, -0.619237, -2.806740, -1.286411, 1.570796, 1.873970],accel_mss,speed_ms,0,blend_radius_m)
  speed_ms = 0.005
  movel([0.303174, -0.624988, -2.813527, -1.273874, 1.570796, 1.873970],accel_mss,speed_ms,0,blend_radius_m)
  speed_ms = 0.025
  movel([0.308567, -0.613243, -2.814565, -1.284581, 1.570796, 1.879363],accel_mss,speed_ms,0,blend_radius_m)
  movel([0.311017, -0.608256, -2.814988, -1.289144, 1.570796, 1.881813],accel_mss,speed_ms,0,blend_radius_m)
  movel([0.313262, -0.603325, -2.815398, -1.293666, 1.570796, 1.884058],accel_mss,speed_ms,0,blend_radius_m)
  movel([0.314771, -0.599239, -2.815730, -1.297420, 1.570796, 1.885567],accel_mss,speed_ms,0,blend_radius_m)
  movel([0.315798, -0.595414, -2.816035, -1.300940, 1.570796, 1.886594],accel_mss,speed_ms,0,blend_radius_m)
  movel([0.316319, -0.591929, -2.816307, -1.304153, 1.570796, 1.887116],accel_mss,speed_ms,0,blend_radius_m)
  movel([0.316316, -0.588864, -2.816543, -1.306981, 1.570796, 1.887112],accel_mss,speed_ms,0,blend_radius_m)
  movel([0.318007, -0.587553, -2.816643, -1.308193, 1.570796, 1.888803],accel_mss,speed_ms,0,blend_radius_m)
  movel([0.319623, -0.586636, -2.816713, -1.309040, 1.570796, 1.890419],accel_mss,speed_ms,0,blend_radius_m)
  movel([0.322733, -0.585300, -2.816813, -1.310275, 1.570796, 1.893529],accel_mss,speed_ms,0,blend_radius_m)
  movel([0.326035, -0.583602, -2.816940, -1.311847, 1.570796, 1.896831],accel_mss,speed_ms,0,blend_radius_m)
  movel([0.327738, -0.582327, -2.817035, -1.313027, 1.570796, 1.898535],accel_mss,speed_ms,0,blend_radius_m)
  movel([0.329386, -0.580626, -2.817160, -1.314604, 1.570796, 1.900182],accel_mss,speed_ms,0,blend_radius_m)
  movel([0.348272, -0.558085, -2.818714, -1.335589, 1.570796, 1.919069],accel_mss,speed_ms,0,blend_radius_m)
  movel([0.348583, -0.555681, -2.818869, -1.337839, 1.570796, 1.919380],accel_mss,speed_ms,0,blend_radius_m)
  movel([0.348124, -0.553879, -2.818983, -1.339527, 1.570796, 1.918921],accel_mss,speed_ms,0,blend_radius_m)
  movel([0.346919, -0.552774, -2.819053, -1.340562, 1.570796, 1.917716],accel_mss,speed_ms,0,blend_radius_m)
  movel([0.345019, -0.552447, -2.819073, -1.340869, 1.570796, 1.915815],accel_mss,speed_ms,0,blend_radius_m)
  movel([0.348929, -0.550078, -2.819220, -1.343091, 1.570796, 1.919726],accel_mss,speed_ms,0,blend_radius_m)
  movel([0.352511, -0.548521, -2.819316, -1.344552, 1.570796, 1.923308],accel_mss,speed_ms,0,blend_radius_m)
  movel([0.355579, -0.547844, -2.819357, -1.345188, 1.570796, 1.926375],accel_mss,speed_ms,0,blend_radius_m)
  movel([0.357960, -0.548103, -2.819342, -1.344945, 1.570796, 1.928756],accel_mss,speed_ms,0,blend_radius_m)
  speed_ms = 0.005
  movel([0.357960, -0.543646, -2.812439, -1.356304, 1.570796, 1.928756],accel_mss,speed_ms,0,blend_radius_m)
  speed_ms = 0.040
  movel([0.361776, -0.533178, -2.813055, -1.366156, 1.570796, 1.932572],accel_mss,speed_ms,0,blend_radius_m)
  speed_ms = 0.005
  movel([0.361776, -0.537444, -2.819971, -1.354974, 1.570796, 1.932572],accel_mss,speed_ms,0,blend_radius_m)
  speed_ms = 0.025
  movel([0.364576, -0.531477, -2.820305, -1.360607, 1.570796, 1.935373],accel_mss,speed_ms,0,blend_radius_m)
  movel([0.366892, -0.525910, -2.820605, -1.365875, 1.570796, 1.937688],accel_mss,speed_ms,0,blend_radius_m)
  movel([0.368755, -0.520699, -2.820875, -1.370815, 1.570796, 1.939551],accel_mss,speed_ms,0,blend_radius_m)
  movel([0.370195, -0.515803, -2.821120, -1.375466, 1.570796, 1.940991],accel_mss,speed_ms,0,blend_radius_m)
  movel([0.371243, -0.511172, -2.821344, -1.379873, 1.570796, 1.942039],accel_mss,speed_ms,0,blend_radius_m)
  movel([0.371933, -0.506757, -2.821551, -1.384081, 1.570796, 1.942730],accel_mss,speed_ms,0,blend_radius_m)
  movel([0.372379, -0.498384, -2.821923, -1.392082, 1.570796, 1.943176],accel_mss,speed_ms,0,blend_radius_m)
  movel([0.362866, -0.518951, -2.820964, -1.372475, 1.570796, 1.933663],accel_mss,speed_ms,0,blend_radius_m)
  movel([0.363724, -0.516768, -2.821073, -1.374548, 1.570796, 1.934521],accel_mss,speed_ms,0,blend_radius_m)
  movel([0.364223, -0.514805, -2.821169, -1.376415, 1.570796, 1.935019],accel_mss,speed_ms,0,blend_radius_m)
  movel([0.364264, -0.511502, -2.821328, -1.379559, 1.570796, 1.935060],accel_mss,speed_ms,0,blend_radius_m)
  movel([0.363219, -0.508977, -2.821448, -1.381964, 1.570796, 1.934016],accel_mss,speed_ms,0,blend_radius_m)
  movel([0.361350, -0.507155, -2.821532, -1.383702, 1.570796, 1.932147],accel_mss,speed_ms,0,blend_radius_m)
  movel([0.358908, -0.505949, -2.821588, -1.384852, 1.570796, 1.929705],accel_mss,speed_ms,0,blend_radius_m)
  movel([0.356160, -0.505277, -2.821618, -1.385494, 1.570796, 1.926956],accel_mss,speed_ms,0,blend_radius_m)
  movel([0.350805, -0.505160, -2.821623, -1.385606, 1.570796, 1.921601],accel_mss,speed_ms,0,blend_radius_m)
  movel([0.352322, -0.511083, -2.821348, -1.379957, 1.570796, 1.923118],accel_mss,speed_ms,0,blend_radius_m)
  movel([0.352350, -0.514791, -2.821170, -1.376429, 1.570796, 1.923146],accel_mss,speed_ms,0,blend_radius_m)
  movel([0.351411, -0.518984, -2.820962, -1.372443, 1.570796, 1.922207],accel_mss,speed_ms,0,blend_radius_m)
  movel([0.349024, -0.519839, -2.820919, -1.371631, 1.570796, 1.919820],accel_mss,speed_ms,0,blend_radius_m)
  movel([0.346872, -0.520177, -2.820902, -1.371311, 1.570796, 1.917668],accel_mss,speed_ms,0,blend_radius_m)
  movel([0.342914, -0.520000, -2.820911, -1.371479, 1.570796, 1.913711],accel_mss,speed_ms,0,blend_radius_m)
  movel([0.338862, -0.519818, -2.820920, -1.371651, 1.570796, 1.909658],accel_mss,speed_ms,0,blend_radius_m)
  movel([0.336592, -0.520149, -2.820903, -1.371337, 1.570796, 1.907388],accel_mss,speed_ms,0,blend_radius_m)
  movel([0.334061, -0.520975, -2.820861, -1.370553, 1.570796, 1.904857],accel_mss,speed_ms,0,blend_radius_m)
  movel([0.331141, -0.526427, -2.820577, -1.365384, 1.570796, 1.901938],accel_mss,speed_ms,0,blend_radius_m)
  movel([0.329142, -0.531477, -2.820305, -1.360607, 1.570796, 1.899939],accel_mss,speed_ms,0,blend_radius_m)
  movel([0.325579, -0.533110, -2.820215, -1.359064, 1.570796, 1.896375],accel_mss,speed_ms,0,blend_radius_m)
  movel([0.322366, -0.534043, -2.820163, -1.358183, 1.570796, 1.893163],accel_mss,speed_ms,0,blend_radius_m)
  movel([0.319565, -0.534258, -2.820151, -1.357980, 1.570796, 1.890361],accel_mss,speed_ms,0,blend_radius_m)
  movel([0.317254, -0.533747, -2.820179, -1.358462, 1.570796, 1.888051],accel_mss,speed_ms,0,blend_radius_m)
  movel([0.316801, -0.534341, -2.820146, -1.357902, 1.570796, 1.887598],accel_mss,speed_ms,0,blend_radius_m)
  movel([0.312948, -0.541162, -2.819756, -1.351471, 1.570796, 1.883744],accel_mss,speed_ms,0,blend_radius_m)
  movel([0.308518, -0.549539, -2.819254, -1.343596, 1.570796, 1.879314],accel_mss,speed_ms,0,blend_radius_m)
  movel([0.306832, -0.553418, -2.819012, -1.339959, 1.570796, 1.877628],accel_mss,speed_ms,0,blend_radius_m)
  movel([0.305575, -0.556874, -2.818792, -1.336722, 1.570796, 1.876371],accel_mss,speed_ms,0,blend_radius_m)
  movel([0.303731, -0.563644, -2.818349, -1.330396, 1.570796, 1.874527],accel_mss,speed_ms,0,blend_radius_m)
  movel([0.296179, -0.560319, -2.818569, -1.333501, 1.570796, 1.866975],accel_mss,speed_ms,0,blend_radius_m)
  movel([0.294293, -0.564423, -2.818297, -1.329670, 1.570796, 1.865090],accel_mss,speed_ms,0,blend_radius_m)
  movel([0.292708, -0.568417, -2.818026, -1.325946, 1.570796, 1.863505],accel_mss,speed_ms,0,blend_radius_m)
  movel([0.290333, -0.576043, -2.817491, -1.318854, 1.570796, 1.861129],accel_mss,speed_ms,0,blend_radius_m)
  movel([0.288921, -0.583036, -2.816982, -1.312371, 1.570796, 1.859717],accel_mss,speed_ms,0,blend_radius_m)
  movel([0.288123, -0.591163, -2.816367, -1.304859, 1.570796, 1.858919],accel_mss,speed_ms,0,blend_radius_m)
  movel([0.287779, -0.592250, -2.816282, -1.303856, 1.570796, 1.858575],accel_mss,speed_ms,0,blend_radius_m)
  movel([0.287159, -0.593436, -2.816190, -1.302763, 1.570796, 1.857956],accel_mss,speed_ms,0,blend_radius_m)
  movel([0.285929, -0.595005, -2.816067, -1.301317, 1.570796, 1.856725],accel_mss,speed_ms,0,blend_radius_m)
  movel([0.276804, -0.603865, -2.815353, -1.293171, 1.570796, 1.847600],accel_mss,speed_ms,0,blend_radius_m)
  movel([0.272177, -0.607770, -2.815029, -1.289590, 1.570796, 1.842973],accel_mss,speed_ms,0,blend_radius_m)
  movel([0.270488, -0.608827, -2.814940, -1.288622, 1.570796, 1.841284],accel_mss,speed_ms,0,blend_radius_m)
  movel([0.269521, -0.608931, -2.814932, -1.288527, 1.570796, 1.840317],accel_mss,speed_ms,0,blend_radius_m)
  movel([0.273197, -0.611176, -2.814741, -1.286471, 1.570796, 1.843994],accel_mss,speed_ms,0,blend_radius_m)
  movel([0.275377, -0.611835, -2.814685, -1.285869, 1.570796, 1.846174],accel_mss,speed_ms,0,blend_radius_m)
  movel([0.277763, -0.612189, -2.814655, -1.285545, 1.570796, 1.848560],accel_mss,speed_ms,0,blend_radius_m)
  movel([0.269994, -0.622190, -2.813780, -1.276420, 1.570796, 1.840790],accel_mss,speed_ms,0,blend_radius_m)
  movel([0.261856, -0.633174, -2.812772, -1.266443, 1.570796, 1.832652],accel_mss,speed_ms,0,blend_radius_m)
  movel([0.258032, -0.638709, -2.812245, -1.261435, 1.570796, 1.828829],accel_mss,speed_ms,0,blend_radius_m)
  movel([0.254566, -0.644093, -2.811721, -1.256575, 1.570796, 1.825362],accel_mss,speed_ms,0,blend_radius_m)
  movel([0.251604, -0.649211, -2.811212, -1.251966, 1.570796, 1.822400],accel_mss,speed_ms,0,blend_radius_m)
  movel([0.249284, -0.653934, -2.810732, -1.247723, 1.570796, 1.820080],accel_mss,speed_ms,0,blend_radius_m)
  movel([0.252859, -0.650213, -2.811111, -1.251065, 1.570796, 1.823656],accel_mss,speed_ms,0,blend_radius_m)
  movel([0.256515, -0.646782, -2.811455, -1.254152, 1.570796, 1.827311],accel_mss,speed_ms,0,blend_radius_m)
  movel([0.260205, -0.643717, -2.811758, -1.256914, 1.570796, 1.831001],accel_mss,speed_ms,0,blend_radius_m)
  movel([0.263905, -0.641082, -2.812016, -1.259292, 1.570796, 1.834702],accel_mss,speed_ms,0,blend_radius_m)
  movel([0.261399, -0.644076, -2.811723, -1.256590, 1.570796, 1.832196],accel_mss,speed_ms,0,blend_radius_m)
  movel([0.256818, -0.650292, -2.811103, -1.250994, 1.570796, 1.827614],accel_mss,speed_ms,0,blend_radius_m)
  movel([0.254774, -0.653463, -2.810780, -1.248146, 1.570796, 1.825570],accel_mss,speed_ms,0,blend_radius_m)
  movel([0.251273, -0.659752, -2.810128, -1.242508, 1.570796, 1.822070],accel_mss,speed_ms,0,blend_radius_m)
  movel([0.249845, -0.662824, -2.809804, -1.239761, 1.570796, 1.820641],accel_mss,speed_ms,0,blend_radius_m)
  movel([0.248659, -0.665801, -2.809486, -1.237103, 1.570796, 1.819455],accel_mss,speed_ms,0,blend_radius_m)
  speed_ms = 0.005
  movel([0.248659, -0.659427, -2.802776, -1.250186, 1.570796, 1.819455],accel_mss,speed_ms,0,blend_radius_m)
  speed_ms = 0.040
  movel([0.261096, -0.660613, -2.802649, -1.249127, 1.570796, 1.831893],accel_mss,speed_ms,0,blend_radius_m)
  speed_ms = 0.005
  movel([0.261096, -0.667004, -2.809356, -1.236029, 1.570796, 1.831893],accel_mss,speed_ms,0,blend_radius_m)
  speed_ms = 0.025
  movel([0.261978, -0.663267, -2.809757, -1.239365, 1.570796, 1.832775],accel_mss,speed_ms,0,blend_radius_m)
  movel([0.263180, -0.659309, -2.810175, -1.242906, 1.570796, 1.833976],accel_mss,speed_ms,0,blend_radius_m)
  movel([0.264694, -0.655166, -2.810606, -1.246618, 1.570796, 1.835491],accel_mss,speed_ms,0,blend_radius_m)
  movel([0.266514, -0.650881, -2.811043, -1.250465, 1.570796, 1.837310],accel_mss,speed_ms,0,blend_radius_m)
  movel([0.268640, -0.646485, -2.811484, -1.254420, 1.570796, 1.839436],accel_mss,speed_ms,0,blend_radius_m)
  movel([0.271058, -0.642019, -2.811924, -1.258445, 1.570796, 1.841854],accel_mss,speed_ms,0,blend_radius_m)
  movel([0.273763, -0.637518, -2.812360, -1.262511, 1.570796, 1.844560],accel_mss,speed_ms,0,blend_radius_m)
  movel([0.276750, -0.633027, -2.812786, -1.266577, 1.570796, 1.847547],accel_mss,speed_ms,0,blend_radius_m)
  movel([0.286612, -0.619041, -2.814060, -1.279289, 1.570796, 1.857408],accel_mss,speed_ms,0,blend_radius_m)
  movel([0.288661, -0.615766, -2.814347, -1.282277, 1.570796, 1.859457],accel_mss,speed_ms,0,blend_radius_m)
  movel([0.290516, -0.612415, -2.814636, -1.285338, 1.570796, 1.861312],accel_mss,speed_ms,0,blend_radius_m)
  movel([0.292163, -0.608913, -2.814933, -1.288542, 1.570796, 1.862959],accel_mss,speed_ms,0,blend_radius_m)
  movel([0.293595, -0.605168, -2.815246, -1.291975, 1.570796, 1.864391],accel_mss,speed_ms,0,blend_radius_m)
  movel([0.296721, -0.594813, -2.816082, -1.301494, 1.570796, 1.867517],accel_mss,speed_ms,0,blend_radius_m)
  movel([0.298529, -0.589512, -2.816494, -1.306384, 1.570796, 1.869326],accel_mss,speed_ms,0,blend_radius_m)
  movel([0.301036, -0.583879, -2.816920, -1.311591, 1.570796, 1.871832],accel_mss,speed_ms,0,blend_radius_m)
  movel([0.303004, -0.580321, -2.817182, -1.314886, 1.570796, 1.873800],accel_mss,speed_ms,0,blend_radius_m)
  movel([0.305252, -0.576741, -2.817442, -1.318207, 1.570796, 1.876048],accel_mss,speed_ms,0,blend_radius_m)
  movel([0.310421, -0.569568, -2.817946, -1.324874, 1.570796, 1.881218],accel_mss,speed_ms,0,blend_radius_m)
  movel([0.316191, -0.562440, -2.818429, -1.331520, 1.570796, 1.886988],accel_mss,speed_ms,0,blend_radius_m)
  movel([0.322221, -0.555435, -2.818884, -1.338070, 1.570796, 1.893018],accel_mss,speed_ms,0,blend_radius_m)
  movel([0.328174, -0.548743, -2.819302, -1.344343, 1.570796, 1.898970],accel_mss,speed_ms,0,blend_radius_m)
  movel([0.334338, -0.542331, -2.819687, -1.350370, 1.570796, 1.905134],accel_mss,speed_ms,0,blend_radius_m)
  movel([0.337426, -0.539436, -2.819856, -1.353096, 1.570796, 1.908222],accel_mss,speed_ms,0,blend_radius_m)
  movel([0.340487, -0.536847, -2.820005, -1.355538, 1.570796, 1.911284],accel_mss,speed_ms,0,blend_radius_m)
  movel([0.343472, -0.534665, -2.820128, -1.357596, 1.570796, 1.914269],accel_mss,speed_ms,0,blend_radius_m)
  movel([0.346372, -0.532952, -2.820223, -1.359214, 1.570796, 1.917168],accel_mss,speed_ms,0,blend_radius_m)
  speed_ms = 0.005
  movel([0.346372, -0.528766, -2.813303, -1.370320, 1.570796, 1.917168],accel_mss,speed_ms,0,blend_radius_m)
  speed_ms = 0.040
  movel([0.349211, -0.530245, -2.813220, -1.368924, 1.570796, 1.920007],accel_mss,speed_ms,0,blend_radius_m)
  speed_ms = 0.005
  movel([0.349211, -0.534458, -2.820140, -1.357792, 1.570796, 1.920007],accel_mss,speed_ms,0,blend_radius_m)
  speed_ms = 0.025
  movel([0.350136, -0.534788, -2.820121, -1.357480, 1.570796, 1.920932],accel_mss,speed_ms,0,blend_radius_m)
  movel([0.351314, -0.535555, -2.820078, -1.356757, 1.570796, 1.922110],accel_mss,speed_ms,0,blend_radius_m)
  movel([0.352745, -0.538693, -2.819899, -1.353797, 1.570796, 1.923541],accel_mss,speed_ms,0,blend_radius_m)
  movel([0.352995, -0.540751, -2.819780, -1.351858, 1.570796, 1.923791],accel_mss,speed_ms,0,blend_radius_m)
  movel([0.352756, -0.541999, -2.819707, -1.350683, 1.570796, 1.923552],accel_mss,speed_ms,0,blend_radius_m)
  movel([0.352424, -0.542400, -2.819683, -1.350305, 1.570796, 1.923220],accel_mss,speed_ms,0,blend_radius_m)
  movel([0.351896, -0.542553, -2.819674, -1.350161, 1.570796, 1.922692],accel_mss,speed_ms,0,blend_radius_m)
  movel([0.346949, -0.542252, -2.819692, -1.350445, 1.570796, 1.917745],accel_mss,speed_ms,0,blend_radius_m)
  movel([0.344047, -0.542790, -2.819660, -1.349939, 1.570796, 1.914843],accel_mss,speed_ms,0,blend_radius_m)
  movel([0.342393, -0.543507, -2.819618, -1.349264, 1.570796, 1.913189],accel_mss,speed_ms,0,blend_radius_m)
  movel([0.340568, -0.544612, -2.819552, -1.348225, 1.570796, 1.911364],accel_mss,speed_ms,0,blend_radius_m)
  movel([0.338416, -0.546316, -2.819450, -1.346623, 1.570796, 1.909212],accel_mss,speed_ms,0,blend_radius_m)
  movel([0.336248, -0.548307, -2.819329, -1.344752, 1.570796, 1.907045],accel_mss,speed_ms,0,blend_radius_m)
  movel([0.330981, -0.553604, -2.819000, -1.339784, 1.570796, 1.901778],accel_mss,speed_ms,0,blend_radius_m)
  movel([0.325797, -0.559304, -2.818635, -1.334450, 1.570796, 1.896593],accel_mss,speed_ms,0,blend_radius_m)
  movel([0.320854, -0.565226, -2.818243, -1.328921, 1.570796, 1.891650],accel_mss,speed_ms,0,blend_radius_m)
  movel([0.316321, -0.571166, -2.817836, -1.323387, 1.570796, 1.887118],accel_mss,speed_ms,0,blend_radius_m)
  movel([0.318210, -0.575456, -2.817533, -1.319400, 1.570796, 1.889007],accel_mss,speed_ms,0,blend_radius_m)
  movel([0.319268, -0.580580, -2.817163, -1.314646, 1.570796, 1.890065],accel_mss,speed_ms,0,blend_radius_m)
  movel([0.317463, -0.580345, -2.817180, -1.314864, 1.570796, 1.888260],accel_mss,speed_ms,0,blend_radius_m)
  movel([0.315279, -0.580728, -2.817152, -1.314509, 1.570796, 1.886076],accel_mss,speed_ms,0,blend_radius_m)
  movel([0.312783, -0.581727, -2.817079, -1.313583, 1.570796, 1.883579],accel_mss,speed_ms,0,blend_radius_m)
  movel([0.310067, -0.583299, -2.816963, -1.312127, 1.570796, 1.880864],accel_mss,speed_ms,0,blend_radius_m)
  movel([0.308732, -0.584478, -2.816875, -1.311036, 1.570796, 1.879528],accel_mss,speed_ms,0,blend_radius_m)
  movel([0.308074, -0.585811, -2.816775, -1.309803, 1.570796, 1.878870],accel_mss,speed_ms,0,blend_radius_m)
  movel([0.303568, -0.599203, -2.815733, -1.297453, 1.570796, 1.874364],accel_mss,speed_ms,0,blend_radius_m)
  movel([0.300842, -0.606188, -2.815161, -1.291040, 1.570796, 1.871639],accel_mss,speed_ms,0,blend_radius_m)
  movel([0.297673, -0.613430, -2.814549, -1.284410, 1.570796, 1.868470],accel_mss,speed_ms,0,blend_radius_m)
  movel([0.294091, -0.620752, -2.813908, -1.277729, 1.570796, 1.864887],accel_mss,speed_ms,0,blend_radius_m)
  movel([0.290108, -0.627994, -2.813253, -1.271142, 1.570796, 1.860904],accel_mss,speed_ms,0,blend_radius_m)
  movel([0.281824, -0.642491, -2.811878, -1.258020, 1.570796, 1.852621],accel_mss,speed_ms,0,blend_radius_m)
  movel([0.278355, -0.649475, -2.811185, -1.251729, 1.570796, 1.849151],accel_mss,speed_ms,0,blend_radius_m)
  movel([0.275692, -0.656248, -2.810494, -1.245647, 1.570796, 1.846488],accel_mss,speed_ms,0,blend_radius_m)
  speed_ms = 0.005
  movel([0.275692, -0.650016, -2.803765, -1.258608, 1.570796, 1.846488],accel_mss,speed_ms,0,blend_radius_m)
  speed_ms = 0.040
  movel([0.303078, -0.630459, -2.805701, -1.276229, 1.570796, 1.873874],accel_mss,speed_ms,0,blend_radius_m)
  speed_ms = 0.005
  movel([0.303078, -0.636388, -2.812468, -1.263533, 1.570796, 1.873874],accel_mss,speed_ms,0,blend_radius_m)
  speed_ms = 0.025
  movel([0.300877, -0.641931, -2.811933, -1.258525, 1.570796, 1.871673],accel_mss,speed_ms,0,blend_radius_m)
  movel([0.297944, -0.647697, -2.811364, -1.253328, 1.570796, 1.868740],accel_mss,speed_ms,0,blend_radius_m)
  movel([0.294388, -0.653488, -2.810778, -1.248123, 1.570796, 1.865184],accel_mss,speed_ms,0,blend_radius_m)
  movel([0.290325, -0.659120, -2.810195, -1.243074, 1.570796, 1.861122],accel_mss,speed_ms,0,blend_radius_m)
  speed_ms = 0.005
  movel([0.290325, -0.652845, -2.803472, -1.256072, 1.570796, 1.861122],accel_mss,speed_ms,0,blend_radius_m)
  speed_ms = 0.040
  movel([0.285559, -0.648924, -2.803877, -1.259587, 1.570796, 1.856356],accel_mss,speed_ms,0,blend_radius_m)
  speed_ms = 0.005
  movel([0.285559, -0.655140, -2.810608, -1.246641, 1.570796, 1.856356],accel_mss,speed_ms,0,blend_radius_m)
  speed_ms = 0.025
  movel([0.265122, -0.690869, -2.806654, -1.214865, 1.570796, 1.835919],accel_mss,speed_ms,0,blend_radius_m)
  movel([0.264110, -0.693065, -2.806393, -1.212930, 1.570796, 1.834906],accel_mss,speed_ms,0,blend_radius_m)
  movel([0.264152, -0.695052, -2.806155, -1.211181, 1.570796, 1.834948],accel_mss,speed_ms,0,blend_radius_m)
  movel([0.264198, -0.697620, -2.805845, -1.208924, 1.570796, 1.834995],accel_mss,speed_ms,0,blend_radius_m)
  movel([0.263580, -0.700665, -2.805474, -1.206250, 1.570796, 1.834376],accel_mss,speed_ms,0,blend_radius_m)
  speed_ms = 0.005
  movel([0.263580, -0.693797, -2.798840, -1.219752, 1.570796, 1.834376],accel_mss,speed_ms,0,blend_radius_m)
  speed_ms = 0.040
  movel([0.294514, -0.667366, -2.801913, -1.243110, 1.570796, 1.865311],accel_mss,speed_ms,0,blend_radius_m)
  speed_ms = 0.005
  movel([0.294514, -0.673858, -2.808605, -1.229926, 1.570796, 1.865311],accel_mss,speed_ms,0,blend_radius_m)
  speed_ms = 0.025
  movel([0.295315, -0.670506, -2.808975, -1.232908, 1.570796, 1.866111],accel_mss,speed_ms,0,blend_radius_m)
  movel([0.296522, -0.666921, -2.809365, -1.236103, 1.570796, 1.867318],accel_mss,speed_ms,0,blend_radius_m)
  movel([0.298113, -0.663163, -2.809768, -1.239458, 1.570796, 1.868909],accel_mss,speed_ms,0,blend_radius_m)
  movel([0.300079, -0.659278, -2.810178, -1.242933, 1.570796, 1.870875],accel_mss,speed_ms,0,blend_radius_m)
  movel([0.301662, -0.656547, -2.810463, -1.245379, 1.570796, 1.872459],accel_mss,speed_ms,0,blend_radius_m)
  movel([0.303456, -0.653817, -2.810744, -1.247828, 1.570796, 1.874252],accel_mss,speed_ms,0,blend_radius_m)
  movel([0.305446, -0.651202, -2.811011, -1.250176, 1.570796, 1.876242],accel_mss,speed_ms,0,blend_radius_m)
  movel([0.307642, -0.648783, -2.811255, -1.252351, 1.570796, 1.878438],accel_mss,speed_ms,0,blend_radius_m)
  movel([0.309571, -0.647096, -2.811424, -1.253869, 1.570796, 1.880367],accel_mss,speed_ms,0,blend_radius_m)
  movel([0.311622, -0.645708, -2.811562, -1.255119, 1.570796, 1.882418],accel_mss,speed_ms,0,blend_radius_m)
  movel([0.313735, -0.644584, -2.811673, -1.256132, 1.570796, 1.884531],accel_mss,speed_ms,0,blend_radius_m)
  movel([0.315866, -0.643684, -2.811761, -1.256943, 1.570796, 1.886662],accel_mss,speed_ms,0,blend_radius_m)
  movel([0.319952, -0.642403, -2.811887, -1.258099, 1.570796, 1.890749],accel_mss,speed_ms,0,blend_radius_m)
  movel([0.323464, -0.641562, -2.811969, -1.258858, 1.570796, 1.894260],accel_mss,speed_ms,0,blend_radius_m)
  movel([0.320966, -0.642401, -2.811887, -1.258101, 1.570796, 1.891763],accel_mss,speed_ms,0,blend_radius_m)
  movel([0.318294, -0.643812, -2.811749, -1.256828, 1.570796, 1.889090],accel_mss,speed_ms,0,blend_radius_m)
  movel([0.315495, -0.645834, -2.811549, -1.255006, 1.570796, 1.886291],accel_mss,speed_ms,0,blend_radius_m)
  movel([0.312607, -0.648515, -2.811282, -1.252592, 1.570796, 1.883404],accel_mss,speed_ms,0,blend_radius_m)
  movel([0.310230, -0.651239, -2.811007, -1.250143, 1.570796, 1.881027],accel_mss,speed_ms,0,blend_radius_m)
  movel([0.308059, -0.654145, -2.810710, -1.247533, 1.570796, 1.878855],accel_mss,speed_ms,0,blend_radius_m)
  movel([0.306173, -0.656981, -2.810418, -1.244991, 1.570796, 1.876970],accel_mss,speed_ms,0,blend_radius_m)
  movel([0.304516, -0.659818, -2.810121, -1.242450, 1.570796, 1.875313],accel_mss,speed_ms,0,blend_radius_m)
  movel([0.301852, -0.665409, -2.809528, -1.237452, 1.570796, 1.872648],accel_mss,speed_ms,0,blend_radius_m)
  movel([0.300013, -0.670719, -2.808951, -1.232718, 1.570796, 1.870810],accel_mss,speed_ms,0,blend_radius_m)
  movel([0.298883, -0.675968, -2.808370, -1.228051, 1.570796, 1.869680],accel_mss,speed_ms,0,blend_radius_m)
  speed_ms = 0.005
  movel([0.298883, -0.669447, -2.801682, -1.241260, 1.570796, 1.869680],accel_mss,speed_ms,0,blend_radius_m)
  speed_ms = 0.040
  movel([0.307826, -0.655875, -2.803154, -1.253360, 1.570796, 1.878622],accel_mss,speed_ms,0,blend_radius_m)
  speed_ms = 0.005
  movel([0.307826, -0.662196, -2.809871, -1.240323, 1.570796, 1.878622],accel_mss,speed_ms,0,blend_radius_m)
  speed_ms = 0.025
  movel([0.307323, -0.663078, -2.809777, -1.239534, 1.570796, 1.878120],accel_mss,speed_ms,0,blend_radius_m)
  movel([0.306534, -0.663658, -2.809715, -1.239016, 1.570796, 1.877330],accel_mss,speed_ms,0,blend_radius_m)
  movel([0.306123, -0.663441, -2.809738, -1.239210, 1.570796, 1.876919],accel_mss,speed_ms,0,blend_radius_m)
  movel([0.306171, -0.662709, -2.809816, -1.239864, 1.570796, 1.876967],accel_mss,speed_ms,0,blend_radius_m)
  movel([0.307220, -0.660803, -2.810018, -1.241568, 1.570796, 1.878017],accel_mss,speed_ms,0,blend_radius_m)
  movel([0.307888, -0.659990, -2.810103, -1.242295, 1.570796, 1.878685],accel_mss,speed_ms,0,blend_radius_m)
  movel([0.308573, -0.659687, -2.810135, -1.242567, 1.570796, 1.879369],accel_mss,speed_ms,0,blend_radius_m)
  movel([0.308862, -0.660078, -2.810094, -1.242217, 1.570796, 1.879658],accel_mss,speed_ms,0,blend_radius_m)
  movel([0.308310, -0.661786, -2.809914, -1.240689, 1.570796, 1.879106],accel_mss,speed_ms,0,blend_radius_m)
  speed_ms = 0.005
  movel([0.308310, -0.655472, -2.803196, -1.253721, 1.570796, 1.879106],accel_mss,speed_ms,0,blend_radius_m)
  speed_ms = 0.040
  movel([0.304559, -0.675854, -2.800959, -1.235576, 1.570796, 1.875355],accel_mss,speed_ms,0,blend_radius_m)
  speed_ms = 0.005
  movel([0.304559, -0.682468, -2.807634, -1.222287, 1.570796, 1.875355],accel_mss,speed_ms,0,blend_radius_m)
  speed_ms = 0.025
  movel([0.307350, -0.678913, -2.808039, -1.225437, 1.570796, 1.878147],accel_mss,speed_ms,0,blend_radius_m)
  movel([0.309763, -0.675323, -2.808442, -1.228624, 1.570796, 1.880560],accel_mss,speed_ms,0,blend_radius_m)
  movel([0.314630, -0.668064, -2.809241, -1.235084, 1.570796, 1.885426],accel_mss,speed_ms,0,blend_radius_m)
  movel([0.318636, -0.663075, -2.809777, -1.239537, 1.570796, 1.889433],accel_mss,speed_ms,0,blend_radius_m)
  movel([0.331896, -0.648234, -2.811310, -1.252845, 1.570796, 1.902692],accel_mss,speed_ms,0,blend_radius_m)
  movel([0.334477, -0.644952, -2.811636, -1.255801, 1.570796, 1.905274],accel_mss,speed_ms,0,blend_radius_m)
  movel([0.335379, -0.643359, -2.811793, -1.257237, 1.570796, 1.906176],accel_mss,speed_ms,0,blend_radius_m)
  movel([0.335707, -0.642027, -2.811924, -1.258439, 1.570796, 1.906504],accel_mss,speed_ms,0,blend_radius_m)
  movel([0.335153, -0.641171, -2.812007, -1.259211, 1.570796, 1.905949],accel_mss,speed_ms,0,blend_radius_m)
  movel([0.333998, -0.641031, -2.812021, -1.259337, 1.570796, 1.904794],accel_mss,speed_ms,0,blend_radius_m)
  movel([0.332045, -0.641265, -2.811998, -1.259126, 1.570796, 1.902842],accel_mss,speed_ms,0,blend_radius_m)
  movel([0.330008, -0.642037, -2.811923, -1.258429, 1.570796, 1.900805],accel_mss,speed_ms,0,blend_radius_m)
  movel([0.327741, -0.643446, -2.811785, -1.257159, 1.570796, 1.898538],accel_mss,speed_ms,0,blend_radius_m)
  movel([0.325107, -0.645580, -2.811574, -1.255234, 1.570796, 1.895903],accel_mss,speed_ms,0,blend_radius_m)
  movel([0.322275, -0.648330, -2.811300, -1.252759, 1.570796, 1.893072],accel_mss,speed_ms,0,blend_radius_m)
  movel([0.319474, -0.651495, -2.810981, -1.249913, 1.570796, 1.890270],accel_mss,speed_ms,0,blend_radius_m)
  movel([0.316738, -0.654946, -2.810628, -1.246815, 1.570796, 1.887534],accel_mss,speed_ms,0,blend_radius_m)
  movel([0.314093, -0.658585, -2.810251, -1.243553, 1.570796, 1.884890],accel_mss,speed_ms,0,blend_radius_m)
  movel([0.309214, -0.665936, -2.809471, -1.236982, 1.570796, 1.880010],accel_mss,speed_ms,0,blend_radius_m)
  movel([0.305058, -0.672658, -2.808738, -1.230993, 1.570796, 1.875854],accel_mss,speed_ms,0,blend_radius_m)
  movel([0.297750, -0.685011, -2.807340, -1.220037, 1.570796, 1.868546],accel_mss,speed_ms,0,blend_radius_m)
  movel([0.295156, -0.689060, -2.806868, -1.216461, 1.570796, 1.865953],accel_mss,speed_ms,0,blend_radius_m)
  movel([0.292310, -0.693059, -2.806394, -1.212936, 1.570796, 1.863107],accel_mss,speed_ms,0,blend_radius_m)
  movel([0.289213, -0.696864, -2.805937, -1.209588, 1.570796, 1.860010],accel_mss,speed_ms,0,blend_radius_m)
  movel([0.285948, -0.700263, -2.805523, -1.206603, 1.570796, 1.856744],accel_mss,speed_ms,0,blend_radius_m)
  movel([0.282594, -0.703051, -2.805179, -1.204158, 1.570796, 1.853391],accel_mss,speed_ms,0,blend_radius_m)
  movel([0.285026, -0.701959, -2.805314, -1.205116, 1.570796, 1.855822],accel_mss,speed_ms,0,blend_radius_m)
  movel([0.287555, -0.700561, -2.805486, -1.206341, 1.570796, 1.858351],accel_mss,speed_ms,0,blend_radius_m)
  movel([0.290159, -0.698865, -2.805694, -1.207830, 1.570796, 1.860956],accel_mss,speed_ms,0,blend_radius_m)
  movel([0.292797, -0.696902, -2.805932, -1.209555, 1.570796, 1.863593],accel_mss,speed_ms,0,blend_radius_m)
  movel([0.292190, -0.699967, -2.805559, -1.206863, 1.570796, 1.862987],accel_mss,speed_ms,0,blend_radius_m)
  movel([0.291131, -0.703283, -2.805151, -1.203956, 1.570796, 1.861928],accel_mss,speed_ms,0,blend_radius_m)
  movel([0.289656, -0.706759, -2.804717, -1.200913, 1.570796, 1.860452],accel_mss,speed_ms,0,blend_radius_m)
  movel([0.287799, -0.710314, -2.804268, -1.197806, 1.570796, 1.858595],accel_mss,speed_ms,0,blend_radius_m)
  movel([0.290896, -0.706539, -2.804745, -1.201105, 1.570796, 1.861693],accel_mss,speed_ms,0,blend_radius_m)
  movel([0.293713, -0.702626, -2.805232, -1.204531, 1.570796, 1.864509],accel_mss,speed_ms,0,blend_radius_m)
  movel([0.296264, -0.698607, -2.805725, -1.208057, 1.570796, 1.867061],accel_mss,speed_ms,0,blend_radius_m)
  movel([0.298581, -0.694511, -2.806220, -1.211658, 1.570796, 1.869377],accel_mss,speed_ms,0,blend_radius_m)
  movel([0.298272, -0.696519, -2.805979, -1.209891, 1.570796, 1.869068],accel_mss,speed_ms,0,blend_radius_m)
  movel([0.297501, -0.698960, -2.805682, -1.207747, 1.570796, 1.868297],accel_mss,speed_ms,0,blend_radius_m)
  movel([0.292554, -0.710490, -2.804246, -1.197653, 1.570796, 1.863350],accel_mss,speed_ms,0,blend_radius_m)
  movel([0.291541, -0.713211, -2.803898, -1.195279, 1.570796, 1.862338],accel_mss,speed_ms,0,blend_radius_m)
  movel([0.290895, -0.715621, -2.803588, -1.193180, 1.570796, 1.861691],accel_mss,speed_ms,0,blend_radius_m)
  movel([0.292970, -0.711559, -2.804110, -1.196720, 1.570796, 1.863766],accel_mss,speed_ms,0,blend_radius_m)
  movel([0.295199, -0.707721, -2.804597, -1.200072, 1.570796, 1.865996],accel_mss,speed_ms,0,blend_radius_m)
  movel([0.300007, -0.700453, -2.805500, -1.206436, 1.570796, 1.870804],accel_mss,speed_ms,0,blend_radius_m)
  movel([0.305109, -0.693243, -2.806372, -1.212774, 1.570796, 1.875905],accel_mss,speed_ms,0,blend_radius_m)
  movel([0.310320, -0.685483, -2.807286, -1.219620, 1.570796, 1.881117],accel_mss,speed_ms,0,blend_radius_m)
  movel([0.313168, -0.680615, -2.807845, -1.223929, 1.570796, 1.883964],accel_mss,speed_ms,0,blend_radius_m)
  movel([0.314986, -0.677889, -2.808154, -1.226346, 1.570796, 1.885783],accel_mss,speed_ms,0,blend_radius_m)
  movel([0.315838, -0.676875, -2.808268, -1.227246, 1.570796, 1.886634],accel_mss,speed_ms,0,blend_radius_m)
  movel([0.316599, -0.676245, -2.808339, -1.227805, 1.570796, 1.887396],accel_mss,speed_ms,0,blend_radius_m)
  movel([0.317214, -0.676071, -2.808359, -1.227960, 1.570796, 1.888010],accel_mss,speed_ms,0,blend_radius_m)
  movel([0.317670, -0.676285, -2.808335, -1.227770, 1.570796, 1.888466],accel_mss,speed_ms,0,blend_radius_m)
  movel([0.318149, -0.677529, -2.808195, -1.226665, 1.570796, 1.888946],accel_mss,speed_ms,0,blend_radius_m)
  movel([0.318083, -0.679329, -2.807992, -1.225069, 1.570796, 1.888880],accel_mss,speed_ms,0,blend_radius_m)
  movel([0.317519, -0.681033, -2.807798, -1.223558, 1.570796, 1.888316],accel_mss,speed_ms,0,blend_radius_m)
  movel([0.320699, -0.674875, -2.808492, -1.229022, 1.570796, 1.891495],accel_mss,speed_ms,0,blend_radius_m)
  movel([0.323397, -0.668795, -2.809162, -1.234432, 1.570796, 1.894193],accel_mss,speed_ms,0,blend_radius_m)
  movel([0.325579, -0.662889, -2.809797, -1.239703, 1.570796, 1.896375],accel_mss,speed_ms,0,blend_radius_m)
  movel([0.327197, -0.657244, -2.810390, -1.244754, 1.570796, 1.897993],accel_mss,speed_ms,0,blend_radius_m)
  speed_ms = 0.005
  movel([0.327197, -0.650997, -2.803664, -1.257728, 1.570796, 1.897993],accel_mss,speed_ms,0,blend_radius_m)
  speed_ms = 0.040
  movel([0.331771, -0.651230, -2.803640, -1.257519, 1.570796, 1.902567],accel_mss,speed_ms,0,blend_radius_m)
  speed_ms = 0.005
  movel([0.331771, -0.657480, -2.810366, -1.244543, 1.570796, 1.902567],accel_mss,speed_ms,0,blend_radius_m)
  speed_ms = 0.025
  movel([0.334530, -0.657298, -2.810385, -1.244706, 1.570796, 1.905327],accel_mss,speed_ms,0,blend_radius_m)
  movel([0.335469, -0.657791, -2.810333, -1.244264, 1.570796, 1.906265],accel_mss,speed_ms,0,blend_radius_m)
  movel([0.335833, -0.658925, -2.810215, -1.243248, 1.570796, 1.906629],accel_mss,speed_ms,0,blend_radius_m)
  movel([0.335591, -0.660382, -2.810062, -1.241945, 1.570796, 1.906388],accel_mss,speed_ms,0,blend_radius_m)
  movel([0.326578, -0.687071, -2.807101, -1.218217, 1.570796, 1.897374],accel_mss,speed_ms,0,blend_radius_m)
  movel([0.325852, -0.688992, -2.806876, -1.216521, 1.570796, 1.896648],accel_mss,speed_ms,0,blend_radius_m)
  movel([0.324885, -0.690983, -2.806641, -1.214765, 1.570796, 1.895681],accel_mss,speed_ms,0,blend_radius_m)
  movel([0.323657, -0.692803, -2.806425, -1.213161, 1.570796, 1.894453],accel_mss,speed_ms,0,blend_radius_m)
  movel([0.322169, -0.694204, -2.806257, -1.211928, 1.570796, 1.892965],accel_mss,speed_ms,0,blend_radius_m)
  movel([0.320845, -0.694805, -2.806185, -1.211399, 1.570796, 1.891642],accel_mss,speed_ms,0,blend_radius_m)
  movel([0.318504, -0.695106, -2.806149, -1.211134, 1.570796, 1.889300],accel_mss,speed_ms,0,blend_radius_m)
  movel([0.317175, -0.695772, -2.806069, -1.210549, 1.570796, 1.887972],accel_mss,speed_ms,0,blend_radius_m)
  movel([0.315504, -0.697448, -2.805866, -1.209075, 1.570796, 1.886301],accel_mss,speed_ms,0,blend_radius_m)
  movel([0.313959, -0.699452, -2.805622, -1.207315, 1.570796, 1.884756],accel_mss,speed_ms,0,blend_radius_m)
  movel([0.312038, -0.701715, -2.805344, -1.205329, 1.570796, 1.882835],accel_mss,speed_ms,0,blend_radius_m)
  movel([0.309999, -0.703714, -2.805097, -1.203577, 1.570796, 1.880795],accel_mss,speed_ms,0,blend_radius_m)
  movel([0.307917, -0.705406, -2.804887, -1.202096, 1.570796, 1.878713],accel_mss,speed_ms,0,blend_radius_m)
  movel([0.305858, -0.706753, -2.804718, -1.200917, 1.570796, 1.876655],accel_mss,speed_ms,0,blend_radius_m)
  movel([0.303892, -0.707720, -2.804597, -1.200072, 1.570796, 1.874689],accel_mss,speed_ms,0,blend_radius_m)
  movel([0.302101, -0.708254, -2.804529, -1.199605, 1.570796, 1.872898],accel_mss,speed_ms,0,blend_radius_m)
  movel([0.300546, -0.708333, -2.804519, -1.199537, 1.570796, 1.871343],accel_mss,speed_ms,0,blend_radius_m)
  movel([0.299304, -0.707895, -2.804575, -1.199919, 1.570796, 1.870100],accel_mss,speed_ms,0,blend_radius_m)
  speed_ms = 0.005
  movel([0.299304, -0.700929, -2.797958, -1.213502, 1.570796, 1.870100],accel_mss,speed_ms,0,blend_radius_m)
  speed_ms = 0.040
  movel([0.281741, -0.727148, -2.794514, -1.190727, 1.570796, 1.852537],accel_mss,speed_ms,0,blend_radius_m)
  speed_ms = 0.005
  movel([0.281741, -0.734459, -2.801067, -1.176863, 1.570796, 1.852537],accel_mss,speed_ms,0,blend_radius_m)
  speed_ms = 0.025
  movel([0.278055, -0.757214, -2.797799, -1.157375, 1.570796, 1.848852],accel_mss,speed_ms,0,blend_radius_m)
  movel([0.277347, -0.760122, -2.797364, -1.154903, 1.570796, 1.848143],accel_mss,speed_ms,0,blend_radius_m)
  movel([0.276648, -0.761640, -2.797135, -1.153614, 1.570796, 1.847444],accel_mss,speed_ms,0,blend_radius_m)
  movel([0.275612, -0.763106, -2.796913, -1.152371, 1.570796, 1.846408],accel_mss,speed_ms,0,blend_radius_m)
  movel([0.272899, -0.765873, -2.796490, -1.150025, 1.570796, 1.843695],accel_mss,speed_ms,0,blend_radius_m)
  movel([0.271996, -0.767514, -2.796238, -1.148637, 1.570796, 1.842792],accel_mss,speed_ms,0,blend_radius_m)
  movel([0.271579, -0.769067, -2.795998, -1.147324, 1.570796, 1.842375],accel_mss,speed_ms,0,blend_radius_m)
  movel([0.271570, -0.771245, -2.795660, -1.145484, 1.570796, 1.842366],accel_mss,speed_ms,0,blend_radius_m)
  movel([0.272150, -0.773015, -2.795383, -1.143991, 1.570796, 1.842946],accel_mss,speed_ms,0,blend_radius_m)
  movel([0.273739, -0.776044, -2.794905, -1.141439, 1.570796, 1.844535],accel_mss,speed_ms,0,blend_radius_m)
  movel([0.274278, -0.778520, -2.794512, -1.139358, 1.570796, 1.845075],accel_mss,speed_ms,0,blend_radius_m)
  movel([0.274468, -0.782488, -2.793874, -1.136027, 1.570796, 1.845264],accel_mss,speed_ms,0,blend_radius_m)
  movel([0.274204, -0.784493, -2.793549, -1.134347, 1.570796, 1.845000],accel_mss,speed_ms,0,blend_radius_m)
  movel([0.273576, -0.786243, -2.793264, -1.132882, 1.570796, 1.844372],accel_mss,speed_ms,0,blend_radius_m)
  movel([0.273096, -0.786948, -2.793148, -1.132292, 1.570796, 1.843892],accel_mss,speed_ms,0,blend_radius_m)
  movel([0.272493, -0.787514, -2.793056, -1.131819, 1.570796, 1.843289],accel_mss,speed_ms,0,blend_radius_m)
  movel([0.271753, -0.787911, -2.792990, -1.131487, 1.570796, 1.842549],accel_mss,speed_ms,0,blend_radius_m)
  movel([0.270866, -0.788109, -2.792958, -1.131322, 1.570796, 1.841663],accel_mss,speed_ms,0,blend_radius_m)
  movel([0.270373, -0.789929, -2.792658, -1.129803, 1.570796, 1.841169],accel_mss,speed_ms,0,blend_radius_m)
  movel([0.270264, -0.791766, -2.792353, -1.128270, 1.570796, 1.841060],accel_mss,speed_ms,0,blend_radius_m)
  movel([0.270864, -0.795336, -2.791756, -1.125297, 1.570796, 1.841661],accel_mss,speed_ms,0,blend_radius_m)
  movel([0.272032, -0.798467, -2.791226, -1.122695, 1.570796, 1.842829],accel_mss,speed_ms,0,blend_radius_m)
  movel([0.273153, -0.800795, -2.790830, -1.120764, 1.570796, 1.843949],accel_mss,speed_ms,0,blend_radius_m)
  movel([0.274846, -0.802928, -2.790464, -1.118997, 1.570796, 1.845642],accel_mss,speed_ms,0,blend_radius_m)
  movel([0.276926, -0.804807, -2.790139, -1.117443, 1.570796, 1.847722],accel_mss,speed_ms,0,blend_radius_m)
  movel([0.278568, -0.807084, -2.789744, -1.115562, 1.570796, 1.849364],accel_mss,speed_ms,0,blend_radius_m)
  movel([0.278969, -0.808565, -2.789485, -1.114339, 1.570796, 1.849766],accel_mss,speed_ms,0,blend_radius_m)
  movel([0.278953, -0.810383, -2.789166, -1.112841, 1.570796, 1.849750],accel_mss,speed_ms,0,blend_radius_m)
  movel([0.278680, -0.811481, -2.788972, -1.111936, 1.570796, 1.849477],accel_mss,speed_ms,0,blend_radius_m)
  movel([0.278145, -0.812669, -2.788762, -1.110959, 1.570796, 1.848941],accel_mss,speed_ms,0,blend_radius_m)
  movel([0.277410, -0.813701, -2.788578, -1.110110, 1.570796, 1.848207],accel_mss,speed_ms,0,blend_radius_m)
  movel([0.276534, -0.814344, -2.788464, -1.109582, 1.570796, 1.847330],accel_mss,speed_ms,0,blend_radius_m)
  movel([0.275921, -0.814398, -2.788454, -1.109537, 1.570796, 1.846718],accel_mss,speed_ms,0,blend_radius_m)
  movel([0.275468, -0.814174, -2.788494, -1.109721, 1.570796, 1.846264],accel_mss,speed_ms,0,blend_radius_m)
  movel([0.271858, -0.811086, -2.789042, -1.112262, 1.570796, 1.842655],accel_mss,speed_ms,0,blend_radius_m)
  movel([0.270330, -0.809207, -2.789372, -1.113809, 1.570796, 1.841127],accel_mss,speed_ms,0,blend_radius_m)
  movel([0.269001, -0.807104, -2.789740, -1.115545, 1.570796, 1.839798],accel_mss,speed_ms,0,blend_radius_m)
  movel([0.268223, -0.808310, -2.789530, -1.114550, 1.570796, 1.839019],accel_mss,speed_ms,0,blend_radius_m)
  movel([0.267662, -0.809516, -2.789318, -1.113555, 1.570796, 1.838458],accel_mss,speed_ms,0,blend_radius_m)
  movel([0.267117, -0.811901, -2.788898, -1.111591, 1.570796, 1.837913],accel_mss,speed_ms,0,blend_radius_m)
  movel([0.267194, -0.814206, -2.788488, -1.109695, 1.570796, 1.837990],accel_mss,speed_ms,0,blend_radius_m)
  movel([0.267740, -0.816372, -2.788101, -1.107916, 1.570796, 1.838537],accel_mss,speed_ms,0,blend_radius_m)
  movel([0.269558, -0.820125, -2.787424, -1.104839, 1.570796, 1.840354],accel_mss,speed_ms,0,blend_radius_m)
  movel([0.271292, -0.822734, -2.786950, -1.102705, 1.570796, 1.842088],accel_mss,speed_ms,0,blend_radius_m)
  movel([0.271782, -0.823852, -2.786745, -1.101792, 1.570796, 1.842578],accel_mss,speed_ms,0,blend_radius_m)
  movel([0.271770, -0.824584, -2.786611, -1.101195, 1.570796, 1.842567],accel_mss,speed_ms,0,blend_radius_m)
  movel([0.271447, -0.825469, -2.786448, -1.100472, 1.570796, 1.842243],accel_mss,speed_ms,0,blend_radius_m)
  movel([0.270811, -0.826430, -2.786271, -1.099689, 1.570796, 1.841608],accel_mss,speed_ms,0,blend_radius_m)
  movel([0.270166, -0.827026, -2.786160, -1.099203, 1.570796, 1.840962],accel_mss,speed_ms,0,blend_radius_m)
  movel([0.268900, -0.827495, -2.786073, -1.098820, 1.570796, 1.839696],accel_mss,speed_ms,0,blend_radius_m)
  movel([0.267192, -0.827915, -2.785996, -1.098478, 1.570796, 1.837988],accel_mss,speed_ms,0,blend_radius_m)
  movel([0.266720, -0.828376, -2.785910, -1.098103, 1.570796, 1.837517],accel_mss,speed_ms,0,blend_radius_m)
  movel([0.266266, -0.829214, -2.785754, -1.097421, 1.570796, 1.837062],accel_mss,speed_ms,0,blend_radius_m)
  movel([0.266043, -0.830090, -2.785591, -1.096708, 1.570796, 1.836840],accel_mss,speed_ms,0,blend_radius_m)
  movel([0.266116, -0.831842, -2.785263, -1.095284, 1.570796, 1.836912],accel_mss,speed_ms,0,blend_radius_m)
  movel([0.266945, -0.834580, -2.784746, -1.093062, 1.570796, 1.837741],accel_mss,speed_ms,0,blend_radius_m)
  movel([0.269138, -0.839974, -2.783718, -1.088697, 1.570796, 1.839934],accel_mss,speed_ms,0,blend_radius_m)
  movel([0.271450, -0.845220, -2.782701, -1.084467, 1.570796, 1.842246],accel_mss,speed_ms,0,blend_radius_m)
  movel([0.271715, -0.846456, -2.782460, -1.083473, 1.570796, 1.842512],accel_mss,speed_ms,0,blend_radius_m)
  movel([0.271667, -0.847931, -2.782170, -1.082288, 1.570796, 1.842463],accel_mss,speed_ms,0,blend_radius_m)
  movel([0.271156, -0.849502, -2.781860, -1.081026, 1.570796, 1.841952],accel_mss,speed_ms,0,blend_radius_m)
  movel([0.270689, -0.850274, -2.781708, -1.080407, 1.570796, 1.841485],accel_mss,speed_ms,0,blend_radius_m)
  movel([0.269378, -0.851585, -2.781448, -1.079356, 1.570796, 1.840175],accel_mss,speed_ms,0,blend_radius_m)
  movel([0.268742, -0.851943, -2.781376, -1.079069, 1.570796, 1.839539],accel_mss,speed_ms,0,blend_radius_m)
  movel([0.267584, -0.852134, -2.781338, -1.078917, 1.570796, 1.838380],accel_mss,speed_ms,0,blend_radius_m)
  movel([0.266607, -0.851814, -2.781402, -1.079173, 1.570796, 1.837403],accel_mss,speed_ms,0,blend_radius_m)
  movel([0.265848, -0.851189, -2.781526, -1.079673, 1.570796, 1.836644],accel_mss,speed_ms,0,blend_radius_m)
  movel([0.262076, -0.846686, -2.782415, -1.083288, 1.570796, 1.832873],accel_mss,speed_ms,0,blend_radius_m)
  movel([0.258644, -0.841774, -2.783371, -1.087244, 1.570796, 1.829441],accel_mss,speed_ms,0,blend_radius_m)
  movel([0.255575, -0.836444, -2.784393, -1.091552, 1.570796, 1.826371],accel_mss,speed_ms,0,blend_radius_m)
  movel([0.252877, -0.830700, -2.785477, -1.096213, 1.570796, 1.823673],accel_mss,speed_ms,0,blend_radius_m)
  movel([0.252039, -0.828406, -2.785904, -1.098078, 1.570796, 1.822835],accel_mss,speed_ms,0,blend_radius_m)
  movel([0.251666, -0.825714, -2.786403, -1.100272, 1.570796, 1.822462],accel_mss,speed_ms,0,blend_radius_m)
  movel([0.251810, -0.823848, -2.786746, -1.101796, 1.570796, 1.822606],accel_mss,speed_ms,0,blend_radius_m)
  movel([0.252185, -0.821837, -2.787113, -1.103439, 1.570796, 1.822981],accel_mss,speed_ms,0,blend_radius_m)
  movel([0.253320, -0.817582, -2.787884, -1.106923, 1.570796, 1.824117],accel_mss,speed_ms,0,blend_radius_m)
  movel([0.258739, -0.801621, -2.790688, -1.120080, 1.570796, 1.829535],accel_mss,speed_ms,0,blend_radius_m)
  movel([0.259950, -0.797210, -2.791440, -1.123739, 1.570796, 1.830746],accel_mss,speed_ms,0,blend_radius_m)
  movel([0.260608, -0.793422, -2.792077, -1.126891, 1.570796, 1.831404],accel_mss,speed_ms,0,blend_radius_m)
  movel([0.260657, -0.791885, -2.792333, -1.128171, 1.570796, 1.831453],accel_mss,speed_ms,0,blend_radius_m)
  movel([0.260469, -0.790661, -2.792536, -1.129192, 1.570796, 1.831265],accel_mss,speed_ms,0,blend_radius_m)
  movel([0.260019, -0.789794, -2.792680, -1.129915, 1.570796, 1.830816],accel_mss,speed_ms,0,blend_radius_m)
  movel([0.259280, -0.789336, -2.792756, -1.130297, 1.570796, 1.830076],accel_mss,speed_ms,0,blend_radius_m)
  movel([0.257564, -0.789210, -2.792776, -1.130402, 1.570796, 1.828361],accel_mss,speed_ms,0,blend_radius_m)
  movel([0.256825, -0.789013, -2.792809, -1.130567, 1.570796, 1.827621],accel_mss,speed_ms,0,blend_radius_m)
  movel([0.256410, -0.788429, -2.792905, -1.131054, 1.570796, 1.827206],accel_mss,speed_ms,0,blend_radius_m)
  movel([0.256635, -0.786836, -2.793167, -1.132386, 1.570796, 1.827431],accel_mss,speed_ms,0,blend_radius_m)
  movel([0.257472, -0.784899, -2.793483, -1.134007, 1.570796, 1.828269],accel_mss,speed_ms,0,blend_radius_m)
  movel([0.260367, -0.778627, -2.794495, -1.139268, 1.570796, 1.831164],accel_mss,speed_ms,0,blend_radius_m)
  movel([0.262974, -0.772428, -2.795475, -1.144486, 1.570796, 1.833770],accel_mss,speed_ms,0,blend_radius_m)
  movel([0.265331, -0.766277, -2.796428, -1.149683, 1.570796, 1.836127],accel_mss,speed_ms,0,blend_radius_m)
  movel([0.267477, -0.760160, -2.797358, -1.154871, 1.570796, 1.838273],accel_mss,speed_ms,0,blend_radius_m)
  movel([0.271335, -0.747950, -2.799160, -1.165279, 1.570796, 1.842131],accel_mss,speed_ms,0,blend_radius_m)
  movel([0.274904, -0.735624, -2.800906, -1.175859, 1.570796, 1.845701],accel_mss,speed_ms,0,blend_radius_m)
  speed_ms = 0.005
  movel([0.274904, -0.728299, -2.794356, -1.189735, 1.570796, 1.845701],accel_mss,speed_ms,0,blend_radius_m)
  speed_ms = 0.040
  movel([0.261432, -0.760067, -2.789732, -1.162590, 1.570796, 1.832228],accel_mss,speed_ms,0,blend_radius_m)
  speed_ms = 0.005
  movel([0.261432, -0.767779, -2.796197, -1.148413, 1.570796, 1.832228],accel_mss,speed_ms,0,blend_radius_m)
  speed_ms = 0.025
  movel([0.254948, -0.776303, -2.794864, -1.141222, 1.570796, 1.825745],accel_mss,speed_ms,0,blend_radius_m)
  movel([0.248348, -0.784582, -2.793535, -1.134272, 1.570796, 1.819145],accel_mss,speed_ms,0,blend_radius_m)
  movel([0.241644, -0.792613, -2.792212, -1.127564, 1.570796, 1.812440],accel_mss,speed_ms,0,blend_radius_m)
  movel([0.234856, -0.800369, -2.790903, -1.121118, 1.570796, 1.805652],accel_mss,speed_ms,0,blend_radius_m)
  movel([0.240164, -0.792420, -2.792244, -1.127725, 1.570796, 1.810961],accel_mss,speed_ms,0,blend_radius_m)
  movel([0.245154, -0.784297, -2.793581, -1.134511, 1.570796, 1.815950],accel_mss,speed_ms,0,blend_radius_m)
  movel([0.249787, -0.776054, -2.794904, -1.141431, 1.570796, 1.820583],accel_mss,speed_ms,0,blend_radius_m)
  movel([0.254028, -0.767747, -2.796202, -1.148440, 1.570796, 1.824825],accel_mss,speed_ms,0,blend_radius_m)
  movel([0.248584, -0.774747, -2.795110, -1.142531, 1.570796, 1.819380],accel_mss,speed_ms,0,blend_radius_m)
  movel([0.243053, -0.781561, -2.794024, -1.136804, 1.570796, 1.813849],accel_mss,speed_ms,0,blend_radius_m)
  movel([0.237436, -0.788187, -2.792945, -1.131257, 1.570796, 1.808232],accel_mss,speed_ms,0,blend_radius_m)
  movel([0.231748, -0.794605, -2.791879, -1.125906, 1.570796, 1.802544],accel_mss,speed_ms,0,blend_radius_m)
  movel([0.225400, -0.801581, -2.790695, -1.120113, 1.570796, 1.796196],accel_mss,speed_ms,0,blend_radius_m)
  movel([0.219321, -0.808709, -2.789460, -1.114220, 1.570796, 1.790117],accel_mss,speed_ms,0,blend_radius_m)
  movel([0.216506, -0.812448, -2.788801, -1.111140, 1.570796, 1.787302],accel_mss,speed_ms,0,blend_radius_m)
  movel([0.213960, -0.816279, -2.788118, -1.107992, 1.570796, 1.784756],accel_mss,speed_ms,0,blend_radius_m)
  movel([0.211819, -0.820113, -2.787427, -1.104849, 1.570796, 1.782615],accel_mss,speed_ms,0,blend_radius_m)
  movel([0.210196, -0.823861, -2.786743, -1.101785, 1.570796, 1.780992],accel_mss,speed_ms,0,blend_radius_m)
  movel([0.211400, -0.819496, -2.787539, -1.105355, 1.570796, 1.782197],accel_mss,speed_ms,0,blend_radius_m)
  movel([0.212956, -0.814870, -2.788370, -1.109149, 1.570796, 1.783752],accel_mss,speed_ms,0,blend_radius_m)
  movel([0.214839, -0.810042, -2.789225, -1.113121, 1.570796, 1.785635],accel_mss,speed_ms,0,blend_radius_m)
  movel([0.217020, -0.805070, -2.790094, -1.117225, 1.570796, 1.787816],accel_mss,speed_ms,0,blend_radius_m)
  movel([0.219468, -0.800018, -2.790963, -1.121409, 1.570796, 1.790265],accel_mss,speed_ms,0,blend_radius_m)
  movel([0.222158, -0.794944, -2.791822, -1.125624, 1.570796, 1.792954],accel_mss,speed_ms,0,blend_radius_m)
  movel([0.225056, -0.789916, -2.792660, -1.129813, 1.570796, 1.795852],accel_mss,speed_ms,0,blend_radius_m)
  movel([0.228128, -0.785006, -2.793466, -1.133918, 1.570796, 1.798924],accel_mss,speed_ms,0,blend_radius_m)
  movel([0.222602, -0.792693, -2.792199, -1.127498, 1.570796, 1.793398],accel_mss,speed_ms,0,blend_radius_m)
  movel([0.217407, -0.800389, -2.790899, -1.121101, 1.570796, 1.788203],accel_mss,speed_ms,0,blend_radius_m)
  movel([0.212522, -0.808071, -2.789571, -1.114747, 1.570796, 1.783318],accel_mss,speed_ms,0,blend_radius_m)
  movel([0.207928, -0.815714, -2.788219, -1.108456, 1.570796, 1.778724],accel_mss,speed_ms,0,blend_radius_m)
  movel([0.203609, -0.823292, -2.786848, -1.102250, 1.570796, 1.774406],accel_mss,speed_ms,0,blend_radius_m)
  movel([0.199541, -0.830784, -2.785461, -1.096144, 1.570796, 1.770338],accel_mss,speed_ms,0,blend_radius_m)
  movel([0.192077, -0.845426, -2.782661, -1.084301, 1.570796, 1.762873],accel_mss,speed_ms,0,blend_radius_m)
  movel([0.194129, -0.840480, -2.783620, -1.088289, 1.570796, 1.764926],accel_mss,speed_ms,0,blend_radius_m)
  movel([0.195772, -0.835299, -2.784610, -1.092480, 1.570796, 1.766568],accel_mss,speed_ms,0,blend_radius_m)
  movel([0.198677, -0.825238, -2.786490, -1.100660, 1.570796, 1.769474],accel_mss,speed_ms,0,blend_radius_m)
  movel([0.200321, -0.820646, -2.787330, -1.104413, 1.570796, 1.771117],accel_mss,speed_ms,0,blend_radius_m)
  movel([0.202086, -0.816428, -2.788091, -1.107870, 1.570796, 1.772882],accel_mss,speed_ms,0,blend_radius_m)
  movel([0.206386, -0.807549, -2.789663, -1.115178, 1.570796, 1.777183],accel_mss,speed_ms,0,blend_radius_m)
  movel([0.205471, -0.808846, -2.789436, -1.114107, 1.570796, 1.776267],accel_mss,speed_ms,0,blend_radius_m)
  movel([0.203922, -0.810541, -2.789138, -1.112710, 1.570796, 1.774718],accel_mss,speed_ms,0,blend_radius_m)
  movel([0.195262, -0.818702, -2.787682, -1.106005, 1.570796, 1.766058],accel_mss,speed_ms,0,blend_radius_m)
  movel([0.192150, -0.821802, -2.787120, -1.103468, 1.570796, 1.762947],accel_mss,speed_ms,0,blend_radius_m)
  movel([0.188692, -0.826170, -2.786318, -1.099900, 1.570796, 1.759489],accel_mss,speed_ms,0,blend_radius_m)
  movel([0.185491, -0.830796, -2.785459, -1.096134, 1.570796, 1.756287],accel_mss,speed_ms,0,blend_radius_m)
  movel([0.179730, -0.840096, -2.783694, -1.088599, 1.570796, 1.750526],accel_mss,speed_ms,0,blend_radius_m)
  movel([0.181985, -0.835282, -2.784614, -1.092494, 1.570796, 1.752782],accel_mss,speed_ms,0,blend_radius_m)
  movel([0.183935, -0.830486, -2.785517, -1.096386, 1.570796, 1.754732],accel_mss,speed_ms,0,blend_radius_m)
  movel([0.187766, -0.820821, -2.787298, -1.104270, 1.570796, 1.758562],accel_mss,speed_ms,0,blend_radius_m)
  movel([0.190156, -0.815689, -2.788224, -1.108477, 1.570796, 1.760953],accel_mss,speed_ms,0,blend_radius_m)
  movel([0.192896, -0.810449, -2.789154, -1.112786, 1.570796, 1.763693],accel_mss,speed_ms,0,blend_radius_m)
  movel([0.199179, -0.799706, -2.791016, -1.121667, 1.570796, 1.769975],accel_mss,speed_ms,0,blend_radius_m)
  movel([0.212906, -0.777998, -2.794595, -1.139796, 1.570796, 1.783702],accel_mss,speed_ms,0,blend_radius_m)
  movel([0.207618, -0.782429, -2.793884, -1.136076, 1.570796, 1.778414],accel_mss,speed_ms,0,blend_radius_m)
  movel([0.202419, -0.787165, -2.793113, -1.132111, 1.570796, 1.773215],accel_mss,speed_ms,0,blend_radius_m)
  movel([0.197333, -0.792166, -2.792286, -1.127937, 1.570796, 1.768130],accel_mss,speed_ms,0,blend_radius_m)
  movel([0.192402, -0.797388, -2.791410, -1.123592, 1.570796, 1.763198],accel_mss,speed_ms,0,blend_radius_m)
  movel([0.187658, -0.802793, -2.790487, -1.119109, 1.570796, 1.758454],accel_mss,speed_ms,0,blend_radius_m)
  movel([0.183125, -0.808351, -2.789522, -1.114516, 1.570796, 1.753921],accel_mss,speed_ms,0,blend_radius_m)
  movel([0.178832, -0.814017, -2.788522, -1.109850, 1.570796, 1.749628],accel_mss,speed_ms,0,blend_radius_m)
  movel([0.174808, -0.819762, -2.787490, -1.105136, 1.570796, 1.745604],accel_mss,speed_ms,0,blend_radius_m)
  movel([0.175871, -0.818014, -2.787806, -1.106569, 1.570796, 1.746668],accel_mss,speed_ms,0,blend_radius_m)
  movel([0.176866, -0.816075, -2.788155, -1.108159, 1.570796, 1.747662],accel_mss,speed_ms,0,blend_radius_m)
  movel([0.178700, -0.811861, -2.788905, -1.111623, 1.570796, 1.749496],accel_mss,speed_ms,0,blend_radius_m)
  movel([0.182052, -0.803765, -2.790319, -1.118305, 1.570796, 1.752849],accel_mss,speed_ms,0,blend_radius_m)
  movel([0.185570, -0.796684, -2.791529, -1.124177, 1.570796, 1.756367],accel_mss,speed_ms,0,blend_radius_m)
  movel([0.189353, -0.789553, -2.792720, -1.130116, 1.570796, 1.760150],accel_mss,speed_ms,0,blend_radius_m)
  movel([0.193392, -0.782376, -2.793892, -1.136121, 1.570796, 1.764188],accel_mss,speed_ms,0,blend_radius_m)
  movel([0.197671, -0.775154, -2.795046, -1.142189, 1.570796, 1.768468],accel_mss,speed_ms,0,blend_radius_m)
  movel([0.202185, -0.767875, -2.796182, -1.148332, 1.570796, 1.772981],accel_mss,speed_ms,0,blend_radius_m)
  movel([0.206927, -0.760544, -2.797300, -1.154544, 1.570796, 1.777723],accel_mss,speed_ms,0,blend_radius_m)
  movel([0.217047, -0.745695, -2.799484, -1.167209, 1.570796, 1.787844],accel_mss,speed_ms,0,blend_radius_m)
  movel([0.212834, -0.750354, -2.798811, -1.163224, 1.570796, 1.783630],accel_mss,speed_ms,0,blend_radius_m)
  movel([0.199928, -0.763515, -2.796851, -1.152024, 1.570796, 1.770724],accel_mss,speed_ms,0,blend_radius_m)
  movel([0.195714, -0.767990, -2.796165, -1.148235, 1.570796, 1.766510],accel_mss,speed_ms,0,blend_radius_m)
  movel([0.191666, -0.772646, -2.795441, -1.144302, 1.570796, 1.762463],accel_mss,speed_ms,0,blend_radius_m)
  movel([0.187933, -0.777464, -2.794680, -1.140245, 1.570796, 1.758729],accel_mss,speed_ms,0,blend_radius_m)
  movel([0.184647, -0.782439, -2.793882, -1.136068, 1.570796, 1.755443],accel_mss,speed_ms,0,blend_radius_m)
  movel([0.189107, -0.774282, -2.795184, -1.142923, 1.570796, 1.759904],accel_mss,speed_ms,0,blend_radius_m)
  movel([0.193566, -0.765777, -2.796505, -1.150107, 1.570796, 1.764363],accel_mss,speed_ms,0,blend_radius_m)
  movel([0.198297, -0.757220, -2.797799, -1.157370, 1.570796, 1.769093],accel_mss,speed_ms,0,blend_radius_m)
  movel([0.200846, -0.753026, -2.798419, -1.160943, 1.570796, 1.771643],accel_mss,speed_ms,0,blend_radius_m)
  movel([0.203569, -0.748941, -2.799016, -1.164432, 1.570796, 1.774365],accel_mss,speed_ms,0,blend_radius_m)
  movel([0.213662, -0.735179, -2.800967, -1.176242, 1.570796, 1.784458],accel_mss,speed_ms,0,blend_radius_m)
  movel([0.224121, -0.721266, -2.802850, -1.188273, 1.570796, 1.794917],accel_mss,speed_ms,0,blend_radius_m)
  movel([0.216555, -0.728535, -2.801877, -1.181977, 1.570796, 1.787351],accel_mss,speed_ms,0,blend_radius_m)
  movel([0.209738, -0.735756, -2.800887, -1.175746, 1.570796, 1.780535],accel_mss,speed_ms,0,blend_radius_m)
  movel([0.203245, -0.743411, -2.799811, -1.169167, 1.570796, 1.774041],accel_mss,speed_ms,0,blend_radius_m)
  movel([0.196669, -0.751954, -2.798577, -1.161858, 1.570796, 1.767465],accel_mss,speed_ms,0,blend_radius_m)
  movel([0.199815, -0.747406, -2.799238, -1.165745, 1.570796, 1.770611],accel_mss,speed_ms,0,blend_radius_m)
  movel([0.202657, -0.742786, -2.799900, -1.169703, 1.570796, 1.773453],accel_mss,speed_ms,0,blend_radius_m)
  movel([0.213090, -0.723806, -2.802513, -1.186070, 1.570796, 1.783886],accel_mss,speed_ms,0,blend_radius_m)
  movel([0.215992, -0.718991, -2.803149, -1.190249, 1.570796, 1.786788],accel_mss,speed_ms,0,blend_radius_m)
  movel([0.219234, -0.714166, -2.803776, -1.194447, 1.570796, 1.790031],accel_mss,speed_ms,0,blend_radius_m)
  movel([0.223935, -0.707979, -2.804564, -1.199846, 1.570796, 1.794731],accel_mss,speed_ms,0,blend_radius_m)
  movel([0.228034, -0.703438, -2.805132, -1.203819, 1.570796, 1.798830],accel_mss,speed_ms,0,blend_radius_m)
  movel([0.228958, -0.702159, -2.805290, -1.204941, 1.570796, 1.799754],accel_mss,speed_ms,0,blend_radius_m)
  movel([0.229281, -0.701076, -2.805423, -1.205890, 1.570796, 1.800078],accel_mss,speed_ms,0,blend_radius_m)
  movel([0.228746, -0.700849, -2.805451, -1.206089, 1.570796, 1.799542],accel_mss,speed_ms,0,blend_radius_m)
  movel([0.227577, -0.701282, -2.805398, -1.205709, 1.570796, 1.798373],accel_mss,speed_ms,0,blend_radius_m)
  movel([0.226000, -0.702187, -2.805286, -1.204915, 1.570796, 1.796796],accel_mss,speed_ms,0,blend_radius_m)
  movel([0.222512, -0.704601, -2.804987, -1.202801, 1.570796, 1.793308],accel_mss,speed_ms,0,blend_radius_m)
  movel([0.220069, -0.706529, -2.804746, -1.201113, 1.570796, 1.790865],accel_mss,speed_ms,0,blend_radius_m)
  movel([0.223947, -0.700924, -2.805442, -1.206023, 1.570796, 1.794743],accel_mss,speed_ms,0,blend_radius_m)
  movel([0.228482, -0.695269, -2.806129, -1.210990, 1.570796, 1.799278],accel_mss,speed_ms,0,blend_radius_m)
  movel([0.237978, -0.684559, -2.807393, -1.220437, 1.570796, 1.808774],accel_mss,speed_ms,0,blend_radius_m)
  speed_ms = 0.005
  movel([0.237978, -0.677915, -2.800723, -1.233751, 1.570796, 1.808774],accel_mss,speed_ms,0,blend_radius_m)
  speed_ms = 0.040
  movel([0.220547, -0.688066, -2.799532, -1.224791, 1.570796, 1.791343],accel_mss,speed_ms,0,blend_radius_m)
  speed_ms = 0.005
  movel([0.220547, -0.694854, -2.806179, -1.211356, 1.570796, 1.791343],accel_mss,speed_ms,0,blend_radius_m)
  speed_ms = 0.025
  movel([0.219117, -0.693473, -2.806345, -1.212571, 1.570796, 1.789913],accel_mss,speed_ms,0,blend_radius_m)
  movel([0.217209, -0.692809, -2.806424, -1.213156, 1.570796, 1.788005],accel_mss,speed_ms,0,blend_radius_m)
  movel([0.214903, -0.692782, -2.806427, -1.213180, 1.570796, 1.785699],accel_mss,speed_ms,0,blend_radius_m)
  movel([0.212279, -0.693307, -2.806365, -1.212717, 1.570796, 1.783076],accel_mss,speed_ms,0,blend_radius_m)
  movel([0.209410, -0.694315, -2.806244, -1.211830, 1.570796, 1.780207],accel_mss,speed_ms,0,blend_radius_m)
  movel([0.206382, -0.695719, -2.806075, -1.210595, 1.570796, 1.777179],accel_mss,speed_ms,0,blend_radius_m)
  movel([0.200145, -0.699383, -2.805631, -1.207376, 1.570796, 1.770941],accel_mss,speed_ms,0,blend_radius_m)
  speed_ms = 0.005
  movel([0.200145, -0.692532, -2.798994, -1.220863, 1.570796, 1.770941],accel_mss,speed_ms,0,blend_radius_m)
  speed_ms = 0.040
  movel([0.225931, -0.670593, -2.801554, -1.240242, 1.570796, 1.796727],accel_mss,speed_ms,0,blend_radius_m)
  speed_ms = 0.005
  movel([0.225931, -0.677131, -2.808240, -1.227018, 1.570796, 1.796727],accel_mss,speed_ms,0,blend_radius_m)
  speed_ms = 0.025
  movel([0.225055, -0.673467, -2.808649, -1.230274, 1.570796, 1.795851],accel_mss,speed_ms,0,blend_radius_m)
  movel([0.223901, -0.670213, -2.809007, -1.233169, 1.570796, 1.794697],accel_mss,speed_ms,0,blend_radius_m)
  movel([0.222358, -0.667526, -2.809299, -1.235564, 1.570796, 1.793155],accel_mss,speed_ms,0,blend_radius_m)
  movel([0.220313, -0.665556, -2.809512, -1.237321, 1.570796, 1.791109],accel_mss,speed_ms,0,blend_radius_m)
  movel([0.217651, -0.664478, -2.809627, -1.238283, 1.570796, 1.788447],accel_mss,speed_ms,0,blend_radius_m)
  movel([0.214276, -0.664423, -2.809633, -1.238332, 1.570796, 1.785072],accel_mss,speed_ms,0,blend_radius_m)
  movel([0.210076, -0.665565, -2.809511, -1.237313, 1.570796, 1.780872],accel_mss,speed_ms,0,blend_radius_m)
  movel([0.207638, -0.666626, -2.809397, -1.236366, 1.570796, 1.778434],accel_mss,speed_ms,0,blend_radius_m)
  movel([0.204957, -0.668041, -2.809244, -1.235104, 1.570796, 1.775753],accel_mss,speed_ms,0,blend_radius_m)
  speed_ms = 0.005
  movel([0.204957, -0.661635, -2.802539, -1.248215, 1.570796, 1.775753],accel_mss,speed_ms,0,blend_radius_m)
  speed_ms = 0.040
  movel([0.226788, -0.643752, -2.804403, -1.264234, 1.570796, 1.797585],accel_mss,speed_ms,0,blend_radius_m)
  speed_ms = 0.005
  movel([0.226788, -0.649888, -2.811144, -1.251357, 1.570796, 1.797585],accel_mss,speed_ms,0,blend_radius_m)
  speed_ms = 0.025
  movel([0.226566, -0.641097, -2.812014, -1.259278, 1.570796, 1.797362],accel_mss,speed_ms,0,blend_radius_m)
  movel([0.225962, -0.637241, -2.812386, -1.262762, 1.570796, 1.796758],accel_mss,speed_ms,0,blend_radius_m)
  movel([0.224859, -0.633949, -2.812699, -1.265741, 1.570796, 1.795656],accel_mss,speed_ms,0,blend_radius_m)
  movel([0.223137, -0.631382, -2.812939, -1.268068, 1.570796, 1.793933],accel_mss,speed_ms,0,blend_radius_m)
  movel([0.220667, -0.629703, -2.813096, -1.269591, 1.570796, 1.791464],accel_mss,speed_ms,0,blend_radius_m)
  movel([0.217324, -0.629062, -2.813155, -1.270172, 1.570796, 1.788120],accel_mss,speed_ms,0,blend_radius_m)
  movel([0.212992, -0.629624, -2.813103, -1.269662, 1.570796, 1.783788],accel_mss,speed_ms,0,blend_radius_m)
  speed_ms = 0.005
  movel([0.212992, -0.623801, -2.806324, -1.282265, 1.570796, 1.783788],accel_mss,speed_ms,0,blend_radius_m)
  speed_ms = 0.040
  movel([0.232327, -0.615376, -2.807086, -1.289927, 1.570796, 1.803124],accel_mss,speed_ms,0,blend_radius_m)
  speed_ms = 0.005
  movel([0.232327, -0.621064, -2.813880, -1.277445, 1.570796, 1.803124],accel_mss,speed_ms,0,blend_radius_m)
  speed_ms = 0.025
  movel([0.233592, -0.614821, -2.814429, -1.283140, 1.570796, 1.804388],accel_mss,speed_ms,0,blend_radius_m)
  movel([0.234489, -0.608705, -2.814951, -1.288733, 1.570796, 1.805285],accel_mss,speed_ms,0,blend_radius_m)
  movel([0.234865, -0.602943, -2.815429, -1.294017, 1.570796, 1.805662],accel_mss,speed_ms,0,blend_radius_m)
  movel([0.234575, -0.597776, -2.815847, -1.298766, 1.570796, 1.805371],accel_mss,speed_ms,0,blend_radius_m)
  movel([0.233465, -0.593433, -2.816190, -1.302766, 1.570796, 1.804261],accel_mss,speed_ms,0,blend_radius_m)
  movel([0.232550, -0.591654, -2.816329, -1.304406, 1.570796, 1.803347],accel_mss,speed_ms,0,blend_radius_m)
  movel([0.229927, -0.589010, -2.816532, -1.306847, 1.570796, 1.800723],accel_mss,speed_ms,0,blend_radius_m)
  movel([0.228177, -0.588212, -2.816593, -1.307584, 1.570796, 1.798973],accel_mss,speed_ms,0,blend_radius_m)
  movel([0.226109, -0.587799, -2.816625, -1.307965, 1.570796, 1.796905],accel_mss,speed_ms,0,blend_radius_m)
  movel([0.223710, -0.587807, -2.816624, -1.307958, 1.570796, 1.794507],accel_mss,speed_ms,0,blend_radius_m)
  speed_ms = 0.005
  movel([0.223710, -0.582664, -2.809776, -1.319949, 1.570796, 1.794507],accel_mss,speed_ms,0,blend_radius_m)
  speed_ms = 0.040
  movel([0.244747, -0.572411, -2.810532, -1.329446, 1.570796, 1.815543],accel_mss,speed_ms,0,blend_radius_m)
  speed_ms = 0.005
  movel([0.244747, -0.577378, -2.817396, -1.317616, 1.570796, 1.815543],accel_mss,speed_ms,0,blend_radius_m)
  speed_ms = 0.025
  movel([0.246755, -0.569725, -2.817936, -1.324728, 1.570796, 1.817551],accel_mss,speed_ms,0,blend_radius_m)
  movel([0.248116, -0.562400, -2.818432, -1.331557, 1.570796, 1.818913],accel_mss,speed_ms,0,blend_radius_m)
  movel([0.248691, -0.555657, -2.818870, -1.337862, 1.570796, 1.819487],accel_mss,speed_ms,0,blend_radius_m)
  movel([0.248301, -0.549791, -2.819238, -1.343360, 1.570796, 1.819097],accel_mss,speed_ms,0,blend_radius_m)
  movel([0.246800, -0.545069, -2.819525, -1.347795, 1.570796, 1.817596],accel_mss,speed_ms,0,blend_radius_m)
  movel([0.245573, -0.543235, -2.819634, -1.349520, 1.570796, 1.816369],accel_mss,speed_ms,0,blend_radius_m)
  movel([0.244017, -0.541784, -2.819720, -1.350886, 1.570796, 1.814813],accel_mss,speed_ms,0,blend_radius_m)
  movel([0.242096, -0.540773, -2.819779, -1.351838, 1.570796, 1.812893],accel_mss,speed_ms,0,blend_radius_m)
  movel([0.239802, -0.540215, -2.819811, -1.352363, 1.570796, 1.810599],accel_mss,speed_ms,0,blend_radius_m)
  movel([0.237118, -0.540162, -2.819814, -1.352413, 1.570796, 1.807915],accel_mss,speed_ms,0,blend_radius_m)
  movel([0.234025, -0.540633, -2.819787, -1.351969, 1.570796, 1.804821],accel_mss,speed_ms,0,blend_radius_m)
  speed_ms = 0.005
  movel([0.234025, -0.536309, -2.812875, -1.363205, 1.570796, 1.804821],accel_mss,speed_ms,0,blend_radius_m)
  speed_ms = 0.040
  movel([0.134268, -0.605369, -2.807954, -1.299066, 1.570796, 1.705065],accel_mss,speed_ms,0,blend_radius_m)
  speed_ms = 0.005
  movel([0.134268, -0.610893, -2.814766, -1.286731, 1.570796, 1.705065],accel_mss,speed_ms,0,blend_radius_m)
  speed_ms = 0.025
  movel([0.139062, -0.610704, -2.814782, -1.286903, 1.570796, 1.709858],accel_mss,speed_ms,0,blend_radius_m)
  movel([0.143343, -0.611341, -2.814727, -1.286320, 1.570796, 1.714139],accel_mss,speed_ms,0,blend_radius_m)
  movel([0.147131, -0.612744, -2.814607, -1.285037, 1.570796, 1.717927],accel_mss,speed_ms,0,blend_radius_m)
  movel([0.150438, -0.614855, -2.814426, -1.283108, 1.570796, 1.721234],accel_mss,speed_ms,0,blend_radius_m)
  movel([0.153266, -0.617622, -2.814184, -1.280583, 1.570796, 1.724062],accel_mss,speed_ms,0,blend_radius_m)
  movel([0.155649, -0.620974, -2.813888, -1.277527, 1.570796, 1.726445],accel_mss,speed_ms,0,blend_radius_m)
  movel([0.157585, -0.624867, -2.813538, -1.273983, 1.570796, 1.728381],accel_mss,speed_ms,0,blend_radius_m)
  movel([0.159113, -0.629220, -2.813140, -1.270029, 1.570796, 1.729909],accel_mss,speed_ms,0,blend_radius_m)
  movel([0.160234, -0.633985, -2.812695, -1.265709, 1.570796, 1.731031],accel_mss,speed_ms,0,blend_radius_m)
  movel([0.160985, -0.639093, -2.812208, -1.261088, 1.570796, 1.731782],accel_mss,speed_ms,0,blend_radius_m)
  movel([0.161377, -0.644483, -2.811683, -1.256224, 1.570796, 1.732173],accel_mss,speed_ms,0,blend_radius_m)
  movel([0.161433, -0.650105, -2.811122, -1.251162, 1.570796, 1.732229],accel_mss,speed_ms,0,blend_radius_m)
  movel([0.161176, -0.655881, -2.810532, -1.245976, 1.570796, 1.731972],accel_mss,speed_ms,0,blend_radius_m)
  movel([0.160617, -0.661779, -2.809915, -1.240696, 1.570796, 1.731414],accel_mss,speed_ms,0,blend_radius_m)
  movel([0.159785, -0.667717, -2.809279, -1.235393, 1.570796, 1.730581],accel_mss,speed_ms,0,blend_radius_m)
  movel([0.158700, -0.673653, -2.808628, -1.230108, 1.570796, 1.729497],accel_mss,speed_ms,0,blend_radius_m)
  movel([0.156908, -0.681704, -2.807721, -1.222964, 1.570796, 1.727704],accel_mss,speed_ms,0,blend_radius_m)
  movel([0.154407, -0.691125, -2.806624, -1.214640, 1.570796, 1.725204],accel_mss,speed_ms,0,blend_radius_m)
  movel([0.151119, -0.701227, -2.805404, -1.205757, 1.570796, 1.721915],accel_mss,speed_ms,0,blend_radius_m)
  movel([0.149156, -0.706325, -2.804772, -1.201292, 1.570796, 1.719952],accel_mss,speed_ms,0,blend_radius_m)
  movel([0.146975, -0.711334, -2.804139, -1.196916, 1.570796, 1.717771],accel_mss,speed_ms,0,blend_radius_m)
  movel([0.144549, -0.716195, -2.803513, -1.192680, 1.570796, 1.715345],accel_mss,speed_ms,0,blend_radius_m)
  movel([0.141880, -0.720809, -2.802910, -1.188670, 1.570796, 1.712676],accel_mss,speed_ms,0,blend_radius_m)
  movel([0.138944, -0.725116, -2.802338, -1.184935, 1.570796, 1.709741],accel_mss,speed_ms,0,blend_radius_m)
  movel([0.135729, -0.729045, -2.801808, -1.181536, 1.570796, 1.706525],accel_mss,speed_ms,0,blend_radius_m)
  movel([0.132223, -0.732511, -2.801335, -1.178542, 1.570796, 1.703020],accel_mss,speed_ms,0,blend_radius_m)
  movel([0.128404, -0.735461, -2.800928, -1.175999, 1.570796, 1.699201],accel_mss,speed_ms,0,blend_radius_m)
  movel([0.126366, -0.736720, -2.800753, -1.174915, 1.570796, 1.697163],accel_mss,speed_ms,0,blend_radius_m)
  movel([0.124243, -0.737826, -2.800599, -1.173964, 1.570796, 1.695039],accel_mss,speed_ms,0,blend_radius_m)
  movel([0.119724, -0.739542, -2.800359, -1.172489, 1.570796, 1.690521],accel_mss,speed_ms,0,blend_radius_m)
  movel([0.114551, -0.740779, -2.800184, -1.171425, 1.570796, 1.685347],accel_mss,speed_ms,0,blend_radius_m)
  movel([0.109817, -0.741377, -2.800100, -1.170912, 1.570796, 1.680614],accel_mss,speed_ms,0,blend_radius_m)
  movel([0.105467, -0.741411, -2.800095, -1.170883, 1.570796, 1.676263],accel_mss,speed_ms,0,blend_radius_m)
  movel([0.101426, -0.740945, -2.800161, -1.171283, 1.570796, 1.672223],accel_mss,speed_ms,0,blend_radius_m)
  movel([0.097644, -0.740044, -2.800288, -1.172057, 1.570796, 1.668440],accel_mss,speed_ms,0,blend_radius_m)
  movel([0.094051, -0.738785, -2.800465, -1.173139, 1.570796, 1.664847],accel_mss,speed_ms,0,blend_radius_m)
  movel([0.087186, -0.735449, -2.800930, -1.176010, 1.570796, 1.657982],accel_mss,speed_ms,0,blend_radius_m)
  movel([0.079841, -0.731436, -2.801483, -1.179470, 1.570796, 1.650638],accel_mss,speed_ms,0,blend_radius_m)
  movel([0.072694, -0.727241, -2.802052, -1.183095, 1.570796, 1.643490],accel_mss,speed_ms,0,blend_radius_m)
  movel([0.065973, -0.722470, -2.802690, -1.187229, 1.570796, 1.636769],accel_mss,speed_ms,0,blend_radius_m)
  movel([0.062851, -0.719732, -2.803052, -1.189606, 1.570796, 1.633647],accel_mss,speed_ms,0,blend_radius_m)
  movel([0.059928, -0.716684, -2.803450, -1.192255, 1.570796, 1.630725],accel_mss,speed_ms,0,blend_radius_m)
  movel([0.056167, -0.713033, -2.803921, -1.195434, 1.570796, 1.626963],accel_mss,speed_ms,0,blend_radius_m)
  movel([0.051841, -0.709928, -2.804317, -1.198143, 1.570796, 1.622637],accel_mss,speed_ms,0,blend_radius_m)
  movel([0.047031, -0.707337, -2.804645, -1.200407, 1.570796, 1.617827],accel_mss,speed_ms,0,blend_radius_m)
  movel([0.041837, -0.705191, -2.804914, -1.202284, 1.570796, 1.612633],accel_mss,speed_ms,0,blend_radius_m)
  movel([0.030653, -0.702051, -2.805303, -1.205035, 1.570796, 1.601450],accel_mss,speed_ms,0,blend_radius_m)
  movel([0.019045, -0.700027, -2.805552, -1.206810, 1.570796, 1.589842],accel_mss,speed_ms,0,blend_radius_m)
  movel([0.009832, -0.699327, -2.805637, -1.207424, 1.570796, 1.580628],accel_mss,speed_ms,0,blend_radius_m)
  movel([-0.000049, -0.699756, -2.805585, -1.207048, 1.570796, 1.570748],accel_mss,speed_ms,0,blend_radius_m)
  movel([-0.010548, -0.701337, -2.805391, -1.205661, 1.570796, 1.560248],accel_mss,speed_ms,0,blend_radius_m)
  movel([-0.021606, -0.704096, -2.805050, -1.203243, 1.570796, 1.549190],accel_mss,speed_ms,0,blend_radius_m)
  movel([-0.033162, -0.708031, -2.804557, -1.199801, 1.570796, 1.537634],accel_mss,speed_ms,0,blend_radius_m)
  movel([-0.039102, -0.710441, -2.804252, -1.197696, 1.570796, 1.531694],accel_mss,speed_ms,0,blend_radius_m)
  movel([-0.051271, -0.716141, -2.803520, -1.192728, 1.570796, 1.519526],accel_mss,speed_ms,0,blend_radius_m)
  movel([-0.057482, -0.719430, -2.803091, -1.189868, 1.570796, 1.513315],accel_mss,speed_ms,0,blend_radius_m)
  movel([-0.070094, -0.726868, -2.802103, -1.183418, 1.570796, 1.500702],accel_mss,speed_ms,0,blend_radius_m)
  movel([-0.078788, -0.732680, -2.801312, -1.178396, 1.570796, 1.492008],accel_mss,speed_ms,0,blend_radius_m)
  movel([-0.087499, -0.739192, -2.800408, -1.172789, 1.570796, 1.483298],accel_mss,speed_ms,0,blend_radius_m)
  movel([-0.096132, -0.746327, -2.799394, -1.166668, 1.570796, 1.474664],accel_mss,speed_ms,0,blend_radius_m)
  movel([-0.104601, -0.754027, -2.798272, -1.160090, 1.570796, 1.466195],accel_mss,speed_ms,0,blend_radius_m)
  movel([-0.112827, -0.762230, -2.797046, -1.153113, 1.570796, 1.457969],accel_mss,speed_ms,0,blend_radius_m)
  movel([-0.120726, -0.770865, -2.795719, -1.145805, 1.570796, 1.450070],accel_mss,speed_ms,0,blend_radius_m)
  movel([-0.128222, -0.779874, -2.794295, -1.138220, 1.570796, 1.442574],accel_mss,speed_ms,0,blend_radius_m)
  movel([-0.135243, -0.789191, -2.792780, -1.130419, 1.570796, 1.435553],accel_mss,speed_ms,0,blend_radius_m)
  movel([-0.141321, -0.798025, -2.791302, -1.123062, 1.570796, 1.429476],accel_mss,speed_ms,0,blend_radius_m)
  movel([-0.146733, -0.806630, -2.789823, -1.115936, 1.570796, 1.424064],accel_mss,speed_ms,0,blend_radius_m)
